Universal Robots URScript: test_first_drawing_7_m18.script

def Machining1():
  # Default parameters:
  global speed_ms = 0.3
  global speed_rads = 0.75
  global accel_mss = 3
  global accel_radss = 1.2
  global blend_radius_m = 0.001

  # Add subprograms here
  # Start of main program
  # Program generated by RoboDK v5.6.5 for UR10e on 02/02/2024 17:08:00
  # Using nominal kinematics.
  blend_radius_m = 0.001
  speed_ms = 1.000
  # set_reference(p[0.133734, -0.230000, -0.017586, 0.000000, 0.000000, 0.000000])
  set_tcp(p[0.000000, 0.000000, 0.252000, 0.000000, 0.000000, 0.000000])
  # Show Tool
  movej([-0.330517, -0.654443, -2.605811, -1.452135, 1.570796, 1.240279],accel_radss,speed_rads,0,blend_radius_m)
  movel([-0.330517, -0.654443, -2.605811, -1.452135, 1.570796, 1.240279],accel_mss,speed_ms,0,blend_radius_m)
  # Splitting Linear movement in 6 (instruction 7: MoveL 3)
  movel([-0.330517, -0.661877, -2.634190, -1.416323, 1.570796, 1.240279],accel_mss,speed_ms,0,blend_radius_m)
  movel([-0.330517, -0.671796, -2.662374, -1.378219, 1.570796, 1.240279],accel_mss,speed_ms,0,blend_radius_m)
  movel([-0.330517, -0.684615, -2.690354, -1.337420, 1.570796, 1.240279],accel_mss,speed_ms,0,blend_radius_m)
  movel([-0.330517, -0.700841, -2.718117, -1.293431, 1.570796, 1.240279],accel_mss,speed_ms,0,blend_radius_m)
  movel([-0.330517, -0.721107, -2.745644, -1.245638, 1.570796, 1.240279],accel_mss,speed_ms,0,blend_radius_m)
  movel([-0.330517, -0.746206, -2.772909, -1.193275, 1.570796, 1.240279],accel_mss,speed_ms,0,blend_radius_m)
  movel([-0.330517, -0.746206, -2.772909, -1.193275, 1.570796, 1.240279],accel_mss,speed_ms,0,blend_radius_m)
  speed_ms = 1.000
  movel([-0.330517, -0.746206, -2.772909, -1.193275, 1.570796, 1.240279],accel_mss,speed_ms,0,blend_radius_m)
  movel([-0.330517, -0.746206, -2.772909, -1.193275, 1.570796, 1.240279],accel_mss,speed_ms,0,blend_radius_m)
  movel([-0.330517, -0.746206, -2.772909, -1.193275, 1.570796, 1.240279],accel_mss,speed_ms,0,blend_radius_m)
  speed_ms = 0.005
  movel([-0.330517, -0.716695, -2.740159, -1.255535, 1.570796, 1.240279],accel_mss,speed_ms,0,blend_radius_m)
  speed_ms = 1.000
  movel([-0.330517, -0.746206, -2.772909, -1.193275, 1.570796, 1.240279],accel_mss,speed_ms,0,blend_radius_m)
  speed_ms = 0.040
  movel([-0.330517, -0.746206, -2.772909, -1.193275, 1.570796, 1.240279],accel_mss,speed_ms,0,blend_radius_m)
  speed_ms = 1.000
  movel([-0.330517, -0.746206, -2.772909, -1.193275, 1.570796, 1.240279],accel_mss,speed_ms,0,blend_radius_m)
  # Splitting Linear movement in 8 (instruction 21: MoveL 12)
  movel([-0.265752, -0.736383, -2.774388, -1.201618, 1.570796, 1.305044],accel_mss,speed_ms,0,blend_radius_m)
  movel([-0.203429, -0.731735, -2.775072, -1.205583, 1.570796, 1.367367],accel_mss,speed_ms,0,blend_radius_m)
  movel([-0.144075, -0.732399, -2.774975, -1.205016, 1.570796, 1.426722],accel_mss,speed_ms,0,blend_radius_m)
  movel([-0.088098, -0.738355, -2.774095, -1.199939, 1.570796, 1.482698],accel_mss,speed_ms,0,blend_radius_m)
  movel([-0.035774, -0.749426, -2.772413, -1.190550, 1.570796, 1.535022],accel_mss,speed_ms,0,blend_radius_m)
  movel([0.012756, -0.765294, -2.769895, -1.177200, 1.570796, 1.583552],accel_mss,speed_ms,0,blend_radius_m)
  movel([0.057475, -0.785519, -2.766498, -1.160372, 1.570796, 1.628271],accel_mss,speed_ms,0,blend_radius_m)
  movel([0.098470, -0.809577, -2.762175, -1.140637, 1.570796, 1.669266],accel_mss,speed_ms,0,blend_radius_m)
  speed_ms = 0.005
  movel([0.098470, -0.850852, -2.793539, -1.067998, 1.570796, 1.669266],accel_mss,speed_ms,0,blend_radius_m)
  speed_ms = 0.025
  movel([0.094484, -0.861595, -2.791431, -1.059363, 1.570796, 1.665281],accel_mss,speed_ms,0,blend_radius_m)
  movel([0.092287, -0.866990, -2.790348, -1.055051, 1.570796, 1.663083],accel_mss,speed_ms,0,blend_radius_m)
  movel([0.089913, -0.872383, -2.789248, -1.050758, 1.570796, 1.660710],accel_mss,speed_ms,0,blend_radius_m)
  movel([0.087338, -0.877755, -2.788135, -1.046499, 1.570796, 1.658135],accel_mss,speed_ms,0,blend_radius_m)
  movel([0.084536, -0.883089, -2.787014, -1.042286, 1.570796, 1.655333],accel_mss,speed_ms,0,blend_radius_m)
  movel([0.081477, -0.888374, -2.785886, -1.038129, 1.570796, 1.652273],accel_mss,speed_ms,0,blend_radius_m)
  movel([0.078131, -0.893592, -2.784756, -1.034042, 1.570796, 1.648928],accel_mss,speed_ms,0,blend_radius_m)
  movel([0.079373, -0.891311, -2.785252, -1.035826, 1.570796, 1.650169],accel_mss,speed_ms,0,blend_radius_m)
  movel([0.080517, -0.888452, -2.785869, -1.038068, 1.570796, 1.651313],accel_mss,speed_ms,0,blend_radius_m)
  movel([0.081210, -0.885772, -2.786443, -1.040174, 1.570796, 1.652007],accel_mss,speed_ms,0,blend_radius_m)
  movel([0.081271, -0.884745, -2.786662, -1.040982, 1.570796, 1.652068],accel_mss,speed_ms,0,blend_radius_m)
  movel([0.081086, -0.884053, -2.786809, -1.041527, 1.570796, 1.651882],accel_mss,speed_ms,0,blend_radius_m)
  movel([0.080605, -0.883776, -2.786868, -1.041745, 1.570796, 1.651401],accel_mss,speed_ms,0,blend_radius_m)
  movel([0.079917, -0.884008, -2.786819, -1.041563, 1.570796, 1.650713],accel_mss,speed_ms,0,blend_radius_m)
  movel([0.079063, -0.884679, -2.786676, -1.041034, 1.570796, 1.649859],accel_mss,speed_ms,0,blend_radius_m)
  movel([0.078060, -0.885737, -2.786451, -1.040201, 1.570796, 1.648856],accel_mss,speed_ms,0,blend_radius_m)
  movel([0.075754, -0.888735, -2.785808, -1.037846, 1.570796, 1.646551],accel_mss,speed_ms,0,blend_radius_m)
  movel([0.073242, -0.892488, -2.784996, -1.034905, 1.570796, 1.644038],accel_mss,speed_ms,0,blend_radius_m)
  movel([0.068514, -0.900288, -2.783281, -1.028820, 1.570796, 1.639311],accel_mss,speed_ms,0,blend_radius_m)
  movel([0.065663, -0.905241, -2.782172, -1.024976, 1.570796, 1.636460],accel_mss,speed_ms,0,blend_radius_m)
  movel([0.061416, -0.912163, -2.780598, -1.019629, 1.570796, 1.632212],accel_mss,speed_ms,0,blend_radius_m)
  movel([0.059067, -0.915476, -2.779833, -1.017080, 1.570796, 1.629863],accel_mss,speed_ms,0,blend_radius_m)
  movel([0.056470, -0.918581, -2.779110, -1.014698, 1.570796, 1.627267],accel_mss,speed_ms,0,blend_radius_m)
  movel([0.057008, -0.917651, -2.779327, -1.015410, 1.570796, 1.627804],accel_mss,speed_ms,0,blend_radius_m)
  movel([0.057386, -0.916311, -2.779639, -1.016439, 1.570796, 1.628182],accel_mss,speed_ms,0,blend_radius_m)
  movel([0.057710, -0.913007, -2.780403, -1.018979, 1.570796, 1.628506],accel_mss,speed_ms,0,blend_radius_m)
  movel([0.057532, -0.909923, -2.781110, -1.021356, 1.570796, 1.628328],accel_mss,speed_ms,0,blend_radius_m)
  movel([0.057276, -0.908855, -2.781354, -1.022180, 1.570796, 1.628072],accel_mss,speed_ms,0,blend_radius_m)
  movel([0.056930, -0.908319, -2.781476, -1.022594, 1.570796, 1.627726],accel_mss,speed_ms,0,blend_radius_m)
  movel([0.055907, -0.908068, -2.781533, -1.022788, 1.570796, 1.626704],accel_mss,speed_ms,0,blend_radius_m)
  movel([0.054873, -0.908367, -2.781465, -1.022557, 1.570796, 1.625669],accel_mss,speed_ms,0,blend_radius_m)
  movel([0.053834, -0.909106, -2.781297, -1.021987, 1.570796, 1.624631],accel_mss,speed_ms,0,blend_radius_m)
  movel([0.052803, -0.910180, -2.781052, -1.021157, 1.570796, 1.623599],accel_mss,speed_ms,0,blend_radius_m)
  movel([0.050825, -0.912852, -2.780439, -1.019098, 1.570796, 1.621621],accel_mss,speed_ms,0,blend_radius_m)
  movel([0.049035, -0.915498, -2.779828, -1.017063, 1.570796, 1.619831],accel_mss,speed_ms,0,blend_radius_m)
  movel([0.046096, -0.919482, -2.778899, -1.014007, 1.570796, 1.616892],accel_mss,speed_ms,0,blend_radius_m)
  movel([0.043104, -0.923120, -2.778043, -1.011226, 1.570796, 1.613900],accel_mss,speed_ms,0,blend_radius_m)
  movel([0.039882, -0.926413, -2.777260, -1.008716, 1.570796, 1.610679],accel_mss,speed_ms,0,blend_radius_m)
  movel([0.036270, -0.929334, -2.776560, -1.006495, 1.570796, 1.607066],accel_mss,speed_ms,0,blend_radius_m)
  movel([0.038295, -0.926302, -2.777286, -1.008800, 1.570796, 1.609092],accel_mss,speed_ms,0,blend_radius_m)
  movel([0.039935, -0.923235, -2.778015, -1.011138, 1.570796, 1.610731],accel_mss,speed_ms,0,blend_radius_m)
  movel([0.040448, -0.921718, -2.778374, -1.012297, 1.570796, 1.611244],accel_mss,speed_ms,0,blend_radius_m)
  movel([0.040644, -0.920343, -2.778697, -1.013349, 1.570796, 1.611440],accel_mss,speed_ms,0,blend_radius_m)
  movel([0.040480, -0.919233, -2.778958, -1.014198, 1.570796, 1.611276],accel_mss,speed_ms,0,blend_radius_m)
  movel([0.039889, -0.918538, -2.779120, -1.014731, 1.570796, 1.610686],accel_mss,speed_ms,0,blend_radius_m)
  movel([0.038611, -0.918412, -2.779150, -1.014827, 1.570796, 1.609407],accel_mss,speed_ms,0,blend_radius_m)
  movel([0.036998, -0.918988, -2.779015, -1.014386, 1.570796, 1.607794],accel_mss,speed_ms,0,blend_radius_m)
  movel([0.035210, -0.920033, -2.778770, -1.013586, 1.570796, 1.606006],accel_mss,speed_ms,0,blend_radius_m)
  movel([0.033415, -0.921289, -2.778475, -1.012625, 1.570796, 1.604211],accel_mss,speed_ms,0,blend_radius_m)
  speed_ms = 0.005
  movel([0.033415, -0.911749, -2.772496, -1.028143, 1.570796, 1.604211],accel_mss,speed_ms,0,blend_radius_m)
  speed_ms = 0.040
  movel([0.037572, -0.944814, -2.764429, -1.003146, 1.570796, 1.608368],accel_mss,speed_ms,0,blend_radius_m)
  speed_ms = 0.005
  movel([0.037572, -0.954534, -2.770284, -0.987571, 1.570796, 1.608368],accel_mss,speed_ms,0,blend_radius_m)
  speed_ms = 0.025
  movel([0.038407, -0.952070, -2.770916, -0.989403, 1.570796, 1.609204],accel_mss,speed_ms,0,blend_radius_m)
  movel([0.039504, -0.949536, -2.771562, -0.991291, 1.570796, 1.610300],accel_mss,speed_ms,0,blend_radius_m)
  movel([0.040832, -0.946976, -2.772211, -0.993202, 1.570796, 1.611628],accel_mss,speed_ms,0,blend_radius_m)
  movel([0.042377, -0.944420, -2.772854, -0.995116, 1.570796, 1.613173],accel_mss,speed_ms,0,blend_radius_m)
  movel([0.044112, -0.941903, -2.773482, -0.997004, 1.570796, 1.614908],accel_mss,speed_ms,0,blend_radius_m)
  movel([0.046017, -0.939467, -2.774087, -0.998835, 1.570796, 1.616813],accel_mss,speed_ms,0,blend_radius_m)
  movel([0.048065, -0.937149, -2.774659, -1.000582, 1.570796, 1.618862],accel_mss,speed_ms,0,blend_radius_m)
  movel([0.050239, -0.934981, -2.775190, -1.002218, 1.570796, 1.621035],accel_mss,speed_ms,0,blend_radius_m)
  movel([0.053602, -0.932102, -2.775891, -1.004396, 1.570796, 1.624398],accel_mss,speed_ms,0,blend_radius_m)
  movel([0.056890, -0.929797, -2.776448, -1.006144, 1.570796, 1.627686],accel_mss,speed_ms,0,blend_radius_m)
  movel([0.060092, -0.928029, -2.776873, -1.007487, 1.570796, 1.630888],accel_mss,speed_ms,0,blend_radius_m)
  movel([0.063188, -0.926767, -2.777175, -1.008446, 1.570796, 1.633984],accel_mss,speed_ms,0,blend_radius_m)
  movel([0.066168, -0.925977, -2.777364, -1.009048, 1.570796, 1.636964],accel_mss,speed_ms,0,blend_radius_m)
  movel([0.069022, -0.925620, -2.777449, -1.009320, 1.570796, 1.639818],accel_mss,speed_ms,0,blend_radius_m)
  movel([0.071734, -0.925666, -2.777438, -1.009285, 1.570796, 1.642530],accel_mss,speed_ms,0,blend_radius_m)
  movel([0.074296, -0.926070, -2.777342, -1.008977, 1.570796, 1.645092],accel_mss,speed_ms,0,blend_radius_m)
  movel([0.076697, -0.926796, -2.777168, -1.008425, 1.570796, 1.647493],accel_mss,speed_ms,0,blend_radius_m)
  movel([0.078931, -0.927802, -2.776927, -1.007659, 1.570796, 1.649727],accel_mss,speed_ms,0,blend_radius_m)
  movel([0.082865, -0.930490, -2.776281, -1.005618, 1.570796, 1.653661],accel_mss,speed_ms,0,blend_radius_m)
  movel([0.086044, -0.933794, -2.775479, -1.003115, 1.570796, 1.656840],accel_mss,speed_ms,0,blend_radius_m)
  movel([0.088410, -0.937397, -2.774597, -1.000394, 1.570796, 1.659206],accel_mss,speed_ms,0,blend_radius_m)
  movel([0.090331, -0.941611, -2.773555, -0.997223, 1.570796, 1.661127],accel_mss,speed_ms,0,blend_radius_m)
  movel([0.091833, -0.946185, -2.772410, -0.993794, 1.570796, 1.662629],accel_mss,speed_ms,0,blend_radius_m)
  movel([0.092966, -0.951056, -2.771175, -0.990158, 1.570796, 1.663762],accel_mss,speed_ms,0,blend_radius_m)
  movel([0.093774, -0.956168, -2.769862, -0.986359, 1.570796, 1.664570],accel_mss,speed_ms,0,blend_radius_m)
  movel([0.094306, -0.961464, -2.768483, -0.982443, 1.570796, 1.665103],accel_mss,speed_ms,0,blend_radius_m)
  movel([0.094614, -0.966887, -2.767050, -0.978453, 1.570796, 1.665411],accel_mss,speed_ms,0,blend_radius_m)
  movel([0.094736, -0.977899, -2.764077, -0.970413, 1.570796, 1.665532],accel_mss,speed_ms,0,blend_radius_m)
  movel([0.094750, -0.985564, -2.761956, -0.964869, 1.570796, 1.665546],accel_mss,speed_ms,0,blend_radius_m)
  movel([0.095064, -0.989150, -2.760950, -0.962290, 1.570796, 1.665861],accel_mss,speed_ms,0,blend_radius_m)
  movel([0.095787, -0.992414, -2.760025, -0.959950, 1.570796, 1.666583],accel_mss,speed_ms,0,blend_radius_m)
  movel([0.097346, -0.996214, -2.758939, -0.957236, 1.570796, 1.668143],accel_mss,speed_ms,0,blend_radius_m)
  movel([0.098905, -1.000023, -2.757839, -0.954527, 1.570796, 1.669701],accel_mss,speed_ms,0,blend_radius_m)
  movel([0.099406, -1.002068, -2.757244, -0.953076, 1.570796, 1.670202],accel_mss,speed_ms,0,blend_radius_m)
  movel([0.099571, -1.004282, -2.756597, -0.951510, 1.570796, 1.670367],accel_mss,speed_ms,0,blend_radius_m)
  movel([0.099295, -1.006711, -2.755882, -0.949796, 1.570796, 1.670091],accel_mss,speed_ms,0,blend_radius_m)
  movel([0.098473, -1.009410, -2.755083, -0.947896, 1.570796, 1.669269],accel_mss,speed_ms,0,blend_radius_m)
  movel([0.101094, -1.002602, -2.757088, -0.952698, 1.570796, 1.671890],accel_mss,speed_ms,0,blend_radius_m)
  movel([0.103419, -0.995838, -2.759047, -0.957504, 1.570796, 1.674215],accel_mss,speed_ms,0,blend_radius_m)
  movel([0.107547, -0.982266, -2.762874, -0.967249, 1.570796, 1.678343],accel_mss,speed_ms,0,blend_radius_m)
  movel([0.109649, -0.974669, -2.764958, -0.972762, 1.570796, 1.680446],accel_mss,speed_ms,0,blend_radius_m)
  movel([0.111578, -0.967069, -2.767001, -0.978319, 1.570796, 1.682375],accel_mss,speed_ms,0,blend_radius_m)
  movel([0.115043, -0.951807, -2.770983, -0.989598, 1.570796, 1.685839],accel_mss,speed_ms,0,blend_radius_m)
  movel([0.118016, -0.936784, -2.774748, -1.000856, 1.570796, 1.688812],accel_mss,speed_ms,0,blend_radius_m)
  movel([0.119175, -0.929313, -2.776564, -1.006511, 1.570796, 1.689972],accel_mss,speed_ms,0,blend_radius_m)
  movel([0.119952, -0.922044, -2.778297, -1.012048, 1.570796, 1.690749],accel_mss,speed_ms,0,blend_radius_m)
  movel([0.120167, -0.916526, -2.779589, -1.016273, 1.570796, 1.690963],accel_mss,speed_ms,0,blend_radius_m)
  movel([0.120127, -0.911118, -2.780837, -1.020434, 1.570796, 1.690923],accel_mss,speed_ms,0,blend_radius_m)
  movel([0.120107, -0.905634, -2.782084, -1.024671, 1.570796, 1.690904],accel_mss,speed_ms,0,blend_radius_m)
  movel([0.120387, -0.899887, -2.783370, -1.029132, 1.570796, 1.691183],accel_mss,speed_ms,0,blend_radius_m)
  movel([0.120647, -0.898247, -2.783733, -1.030409, 1.570796, 1.691443],accel_mss,speed_ms,0,blend_radius_m)
  movel([0.121203, -0.896466, -2.784126, -1.031797, 1.570796, 1.692000],accel_mss,speed_ms,0,blend_radius_m)
  movel([0.122110, -0.894787, -2.784494, -1.033107, 1.570796, 1.692906],accel_mss,speed_ms,0,blend_radius_m)
  movel([0.122719, -0.894054, -2.784655, -1.033680, 1.570796, 1.693515],accel_mss,speed_ms,0,blend_radius_m)
  movel([0.123441, -0.893428, -2.784791, -1.034169, 1.570796, 1.694238],accel_mss,speed_ms,0,blend_radius_m)
  movel([0.124465, -0.892889, -2.784909, -1.034591, 1.570796, 1.695262],accel_mss,speed_ms,0,blend_radius_m)
  movel([0.125422, -0.892628, -2.784965, -1.034795, 1.570796, 1.696219],accel_mss,speed_ms,0,blend_radius_m)
  movel([0.130425, -0.891913, -2.785121, -1.035355, 1.570796, 1.701221],accel_mss,speed_ms,0,blend_radius_m)
  movel([0.134885, -0.891965, -2.785110, -1.035315, 1.570796, 1.705681],accel_mss,speed_ms,0,blend_radius_m)
  movel([0.138838, -0.892713, -2.784947, -1.034729, 1.570796, 1.709634],accel_mss,speed_ms,0,blend_radius_m)
  movel([0.142320, -0.894105, -2.784643, -1.033640, 1.570796, 1.713117],accel_mss,speed_ms,0,blend_radius_m)
  movel([0.145368, -0.896070, -2.784213, -1.032106, 1.570796, 1.716164],accel_mss,speed_ms,0,blend_radius_m)
  movel([0.148021, -0.898542, -2.783668, -1.030179, 1.570796, 1.718817],accel_mss,speed_ms,0,blend_radius_m)
  movel([0.150317, -0.901457, -2.783021, -1.027911, 1.570796, 1.721113],accel_mss,speed_ms,0,blend_radius_m)
  movel([0.152293, -0.904755, -2.782282, -1.025352, 1.570796, 1.723089],accel_mss,speed_ms,0,blend_radius_m)
  movel([0.153993, -0.908367, -2.781465, -1.022557, 1.570796, 1.724789],accel_mss,speed_ms,0,blend_radius_m)
  movel([0.155459, -0.912228, -2.780583, -1.019578, 1.570796, 1.726255],accel_mss,speed_ms,0,blend_radius_m)
  movel([0.157842, -0.920452, -2.778672, -1.013265, 1.570796, 1.728639],accel_mss,speed_ms,0,blend_radius_m)
  movel([0.161526, -0.937276, -2.774627, -1.000486, 1.570796, 1.732322],accel_mss,speed_ms,0,blend_radius_m)
  movel([0.162250, -0.939773, -2.774011, -0.998605, 1.570796, 1.733046],accel_mss,speed_ms,0,blend_radius_m)
  movel([0.162856, -0.940764, -2.773765, -0.997859, 1.570796, 1.733653],accel_mss,speed_ms,0,blend_radius_m)
  movel([0.163731, -0.941443, -2.773597, -0.997349, 1.570796, 1.734527],accel_mss,speed_ms,0,blend_radius_m)
  movel([0.165528, -0.941709, -2.773531, -0.997150, 1.570796, 1.736325],accel_mss,speed_ms,0,blend_radius_m)
  movel([0.166517, -0.941509, -2.773580, -0.997300, 1.570796, 1.737313],accel_mss,speed_ms,0,blend_radius_m)
  movel([0.167553, -0.941108, -2.773680, -0.997601, 1.570796, 1.738350],accel_mss,speed_ms,0,blend_radius_m)
  movel([0.169715, -0.939801, -2.774004, -0.998584, 1.570796, 1.740512],accel_mss,speed_ms,0,blend_radius_m)
  movel([0.171931, -0.937949, -2.774462, -0.999978, 1.570796, 1.742727],accel_mss,speed_ms,0,blend_radius_m)
  movel([0.174106, -0.935721, -2.775009, -1.001659, 1.570796, 1.744902],accel_mss,speed_ms,0,blend_radius_m)
  movel([0.176150, -0.933279, -2.775605, -1.003505, 1.570796, 1.746946],accel_mss,speed_ms,0,blend_radius_m)
  movel([0.177974, -0.930783, -2.776210, -1.005396, 1.570796, 1.748770],accel_mss,speed_ms,0,blend_radius_m)
  movel([0.179471, -0.928409, -2.776782, -1.007198, 1.570796, 1.750268],accel_mss,speed_ms,0,blend_radius_m)
  movel([0.181767, -0.924306, -2.777762, -1.010321, 1.570796, 1.752563],accel_mss,speed_ms,0,blend_radius_m)
  movel([0.183931, -0.920150, -2.778743, -1.013496, 1.570796, 1.754728],accel_mss,speed_ms,0,blend_radius_m)
  movel([0.187846, -0.911748, -2.780693, -1.019948, 1.570796, 1.758643],accel_mss,speed_ms,0,blend_radius_m)
  movel([0.191204, -0.903342, -2.782599, -1.026448, 1.570796, 1.762001],accel_mss,speed_ms,0,blend_radius_m)
  movel([0.193979, -0.895073, -2.784432, -1.032884, 1.570796, 1.764775],accel_mss,speed_ms,0,blend_radius_m)
  movel([0.194923, -0.891979, -2.785107, -1.035303, 1.570796, 1.765719],accel_mss,speed_ms,0,blend_radius_m)
  movel([0.196094, -0.888834, -2.785787, -1.037769, 1.570796, 1.766891],accel_mss,speed_ms,0,blend_radius_m)
  movel([0.196862, -0.887263, -2.786124, -1.039002, 1.570796, 1.767658],accel_mss,speed_ms,0,blend_radius_m)
  movel([0.197803, -0.885695, -2.786460, -1.040235, 1.570796, 1.768600],accel_mss,speed_ms,0,blend_radius_m)
  movel([0.198955, -0.884142, -2.786790, -1.041457, 1.570796, 1.769752],accel_mss,speed_ms,0,blend_radius_m)
  movel([0.200357, -0.882615, -2.787114, -1.042660, 1.570796, 1.771153],accel_mss,speed_ms,0,blend_radius_m)
  movel([0.202401, -0.881008, -2.787453, -1.043928, 1.570796, 1.773197],accel_mss,speed_ms,0,blend_radius_m)
  movel([0.204401, -0.880128, -2.787638, -1.044623, 1.570796, 1.775198],accel_mss,speed_ms,0,blend_radius_m)
  movel([0.206224, -0.879892, -2.787688, -1.044809, 1.570796, 1.777021],accel_mss,speed_ms,0,blend_radius_m)
  movel([0.207752, -0.880207, -2.787622, -1.044560, 1.570796, 1.778548],accel_mss,speed_ms,0,blend_radius_m)
  movel([0.209849, -0.881389, -2.787373, -1.043627, 1.570796, 1.780645],accel_mss,speed_ms,0,blend_radius_m)
  movel([0.211668, -0.882983, -2.787036, -1.042370, 1.570796, 1.782464],accel_mss,speed_ms,0,blend_radius_m)
  movel([0.214678, -0.886847, -2.786213, -1.039329, 1.570796, 1.785474],accel_mss,speed_ms,0,blend_radius_m)
  movel([0.215840, -0.888920, -2.785768, -1.037701, 1.570796, 1.786637],accel_mss,speed_ms,0,blend_radius_m)
  movel([0.216722, -0.891180, -2.785280, -1.035929, 1.570796, 1.787518],accel_mss,speed_ms,0,blend_radius_m)
  movel([0.217344, -0.893608, -2.784752, -1.034029, 1.570796, 1.788140],accel_mss,speed_ms,0,blend_radius_m)
  movel([0.217717, -0.896195, -2.784185, -1.032008, 1.570796, 1.788513],accel_mss,speed_ms,0,blend_radius_m)
  movel([0.217858, -0.898923, -2.783584, -1.029882, 1.570796, 1.788654],accel_mss,speed_ms,0,blend_radius_m)
  movel([0.217499, -0.904763, -2.782280, -1.025346, 1.570796, 1.788295],accel_mss,speed_ms,0,blend_radius_m)
  movel([0.217027, -0.907846, -2.781583, -1.022960, 1.570796, 1.787823],accel_mss,speed_ms,0,blend_radius_m)
  movel([0.215585, -0.914270, -2.780112, -1.018007, 1.570796, 1.786381],accel_mss,speed_ms,0,blend_radius_m)
  movel([0.213564, -0.920962, -2.778552, -1.012875, 1.570796, 1.784360],accel_mss,speed_ms,0,blend_radius_m)
  movel([0.211074, -0.927836, -2.776919, -1.007633, 1.570796, 1.781870],accel_mss,speed_ms,0,blend_radius_m)
  movel([0.208233, -0.934789, -2.775237, -1.002363, 1.570796, 1.779029],accel_mss,speed_ms,0,blend_radius_m)
  movel([0.203631, -0.944939, -2.772723, -0.994727, 1.570796, 1.774427],accel_mss,speed_ms,0,blend_radius_m)
  movel([0.201108, -0.949995, -2.771446, -0.990948, 1.570796, 1.771904],accel_mss,speed_ms,0,blend_radius_m)
  movel([0.198410, -0.955010, -2.770161, -0.987218, 1.570796, 1.769207],accel_mss,speed_ms,0,blend_radius_m)
  movel([0.195524, -0.959954, -2.768878, -0.983557, 1.570796, 1.766320],accel_mss,speed_ms,0,blend_radius_m)
  movel([0.192436, -0.964804, -2.767603, -0.979982, 1.570796, 1.763232],accel_mss,speed_ms,0,blend_radius_m)
  movel([0.189119, -0.969547, -2.766339, -0.976502, 1.570796, 1.759915],accel_mss,speed_ms,0,blend_radius_m)
  movel([0.185564, -0.974153, -2.765098, -0.973139, 1.570796, 1.756360],accel_mss,speed_ms,0,blend_radius_m)
  movel([0.180277, -0.980341, -2.763406, -0.968642, 1.570796, 1.751073],accel_mss,speed_ms,0,blend_radius_m)
  movel([0.177371, -0.983434, -2.762550, -0.966406, 1.570796, 1.748167],accel_mss,speed_ms,0,blend_radius_m)
  movel([0.174357, -0.986357, -2.761734, -0.964297, 1.570796, 1.745154],accel_mss,speed_ms,0,blend_radius_m)
  movel([0.171294, -0.988986, -2.760996, -0.962407, 1.570796, 1.742090],accel_mss,speed_ms,0,blend_radius_m)
  movel([0.168232, -0.991197, -2.760371, -0.960822, 1.570796, 1.739028],accel_mss,speed_ms,0,blend_radius_m)
  movel([0.165220, -0.992864, -2.759897, -0.959628, 1.570796, 1.736016],accel_mss,speed_ms,0,blend_radius_m)
  movel([0.163750, -0.993460, -2.759727, -0.959202, 1.570796, 1.734546],accel_mss,speed_ms,0,blend_radius_m)
  movel([0.162314, -0.993869, -2.759610, -0.958910, 1.570796, 1.733110],accel_mss,speed_ms,0,blend_radius_m)
  movel([0.160767, -0.994093, -2.759546, -0.958749, 1.570796, 1.731564],accel_mss,speed_ms,0,blend_radius_m)
  movel([0.159366, -0.994058, -2.759556, -0.958774, 1.570796, 1.730163],accel_mss,speed_ms,0,blend_radius_m)
  movel([0.158098, -0.993791, -2.759633, -0.958966, 1.570796, 1.728894],accel_mss,speed_ms,0,blend_radius_m)
  movel([0.156956, -0.993308, -2.759770, -0.959311, 1.570796, 1.727752],accel_mss,speed_ms,0,blend_radius_m)
  movel([0.155007, -0.991802, -2.760199, -0.960388, 1.570796, 1.725804],accel_mss,speed_ms,0,blend_radius_m)
  movel([0.153455, -0.989715, -2.760790, -0.961884, 1.570796, 1.724251],accel_mss,speed_ms,0,blend_radius_m)
  movel([0.152226, -0.987238, -2.761488, -0.963664, 1.570796, 1.723022],accel_mss,speed_ms,0,blend_radius_m)
  movel([0.151254, -0.984552, -2.762239, -0.965599, 1.570796, 1.722051],accel_mss,speed_ms,0,blend_radius_m)
  movel([0.149812, -0.979297, -2.763693, -0.969399, 1.570796, 1.720608],accel_mss,speed_ms,0,blend_radius_m)
  movel([0.149169, -0.976821, -2.764372, -0.971196, 1.570796, 1.719965],accel_mss,speed_ms,0,blend_radius_m)
  movel([0.148254, -0.974605, -2.764975, -0.972809, 1.570796, 1.719050],accel_mss,speed_ms,0,blend_radius_m)
  movel([0.147575, -0.973756, -2.765205, -0.973427, 1.570796, 1.718371],accel_mss,speed_ms,0,blend_radius_m)
  movel([0.146683, -0.973163, -2.765366, -0.973860, 1.570796, 1.717479],accel_mss,speed_ms,0,blend_radius_m)
  movel([0.145535, -0.972893, -2.765439, -0.974057, 1.570796, 1.716332],accel_mss,speed_ms,0,blend_radius_m)
  movel([0.144083, -0.973006, -2.765408, -0.973975, 1.570796, 1.714879],accel_mss,speed_ms,0,blend_radius_m)
  movel([0.144394, -0.973052, -2.765396, -0.973941, 1.570796, 1.715191],accel_mss,speed_ms,0,blend_radius_m)
  movel([0.144561, -0.973335, -2.765319, -0.973734, 1.570796, 1.715357],accel_mss,speed_ms,0,blend_radius_m)
  movel([0.144480, -0.974556, -2.764988, -0.972845, 1.570796, 1.715276],accel_mss,speed_ms,0,blend_radius_m)
  movel([0.143903, -0.976547, -2.764446, -0.971395, 1.570796, 1.714700],accel_mss,speed_ms,0,blend_radius_m)
  movel([0.142911, -0.979182, -2.763725, -0.969482, 1.570796, 1.713708],accel_mss,speed_ms,0,blend_radius_m)
  movel([0.139967, -0.985880, -2.761868, -0.964641, 1.570796, 1.710763],accel_mss,speed_ms,0,blend_radius_m)
  movel([0.136215, -0.993659, -2.759670, -0.959059, 1.570796, 1.707011],accel_mss,speed_ms,0,blend_radius_m)
  movel([0.128486, -1.008701, -2.755293, -0.948395, 1.570796, 1.699282],accel_mss,speed_ms,0,blend_radius_m)
  movel([0.123866, -1.017165, -2.752755, -0.942469, 1.570796, 1.694663],accel_mss,speed_ms,0,blend_radius_m)
  movel([0.118500, -1.025835, -2.750097, -0.936457, 1.570796, 1.689296],accel_mss,speed_ms,0,blend_radius_m)
  movel([0.113088, -1.034273, -2.747454, -0.930662, 1.570796, 1.683885],accel_mss,speed_ms,0,blend_radius_m)
  movel([0.107607, -1.042564, -2.744801, -0.925024, 1.570796, 1.678403],accel_mss,speed_ms,0,blend_radius_m)
  movel([0.096784, -1.058318, -2.739605, -0.914466, 1.570796, 1.667580],accel_mss,speed_ms,0,blend_radius_m)
  movel([0.091340, -1.065635, -2.737121, -0.909633, 1.570796, 1.662136],accel_mss,speed_ms,0,blend_radius_m)
  movel([0.088492, -1.069136, -2.735917, -0.907336, 1.570796, 1.659288],accel_mss,speed_ms,0,blend_radius_m)
  movel([0.085541, -1.072496, -2.734751, -0.905142, 1.570796, 1.656337],accel_mss,speed_ms,0,blend_radius_m)
  movel([0.082458, -1.075684, -2.733635, -0.903069, 1.570796, 1.653255],accel_mss,speed_ms,0,blend_radius_m)
  movel([0.079236, -1.078673, -2.732582, -0.901134, 1.570796, 1.650032],accel_mss,speed_ms,0,blend_radius_m)
  movel([0.080076, -1.072663, -2.734693, -0.905033, 1.570796, 1.650872],accel_mss,speed_ms,0,blend_radius_m)
  movel([0.080087, -1.070990, -2.735275, -0.906125, 1.570796, 1.650884],accel_mss,speed_ms,0,blend_radius_m)
  movel([0.079804, -1.070415, -2.735474, -0.906500, 1.570796, 1.650600],accel_mss,speed_ms,0,blend_radius_m)
  movel([0.079211, -1.070213, -2.735544, -0.906632, 1.570796, 1.650008],accel_mss,speed_ms,0,blend_radius_m)
  movel([0.078545, -1.070393, -2.735482, -0.906514, 1.570796, 1.649341],accel_mss,speed_ms,0,blend_radius_m)
  movel([0.077831, -1.070816, -2.735335, -0.906238, 1.570796, 1.648627],accel_mss,speed_ms,0,blend_radius_m)
  movel([0.074420, -1.073503, -2.734399, -0.904486, 1.570796, 1.645216],accel_mss,speed_ms,0,blend_radius_m)
  movel([0.072411, -1.074760, -2.733960, -0.903669, 1.570796, 1.643207],accel_mss,speed_ms,0,blend_radius_m)
  movel([0.070406, -1.075731, -2.733619, -0.903039, 1.570796, 1.641202],accel_mss,speed_ms,0,blend_radius_m)
  movel([0.068457, -1.076392, -2.733387, -0.902610, 1.570796, 1.639253],accel_mss,speed_ms,0,blend_radius_m)
  movel([0.067876, -1.076424, -2.733376, -0.902590, 1.570796, 1.638673],accel_mss,speed_ms,0,blend_radius_m)
  movel([0.067717, -1.076086, -2.733494, -0.902809, 1.570796, 1.638514],accel_mss,speed_ms,0,blend_radius_m)
  movel([0.068293, -1.074277, -2.734129, -0.903983, 1.570796, 1.639089],accel_mss,speed_ms,0,blend_radius_m)
  movel([0.068248, -1.073755, -2.734312, -0.904323, 1.570796, 1.639044],accel_mss,speed_ms,0,blend_radius_m)
  movel([0.067937, -1.073447, -2.734419, -0.904523, 1.570796, 1.638733],accel_mss,speed_ms,0,blend_radius_m)
  movel([0.067444, -1.073351, -2.734453, -0.904586, 1.570796, 1.638240],accel_mss,speed_ms,0,blend_radius_m)
  movel([0.066848, -1.073466, -2.734412, -0.904511, 1.570796, 1.637644],accel_mss,speed_ms,0,blend_radius_m)
  movel([0.065582, -1.074163, -2.734169, -0.904057, 1.570796, 1.636378],accel_mss,speed_ms,0,blend_radius_m)
  movel([0.056656, -1.081474, -2.731587, -0.899328, 1.570796, 1.627452],accel_mss,speed_ms,0,blend_radius_m)
  movel([0.059293, -1.078836, -2.732524, -0.901029, 1.570796, 1.630089],accel_mss,speed_ms,0,blend_radius_m)
  movel([0.061894, -1.075999, -2.733525, -0.902865, 1.570796, 1.632691],accel_mss,speed_ms,0,blend_radius_m)
  movel([0.064438, -1.073011, -2.734571, -0.904807, 1.570796, 1.635234],accel_mss,speed_ms,0,blend_radius_m)
  movel([0.066915, -1.069903, -2.735651, -0.906834, 1.570796, 1.637712],accel_mss,speed_ms,0,blend_radius_m)
  movel([0.071603, -1.063485, -2.737856, -0.911048, 1.570796, 1.642399],accel_mss,speed_ms,0,blend_radius_m)
  movel([0.075821, -1.057076, -2.740022, -0.915291, 1.570796, 1.646617],accel_mss,speed_ms,0,blend_radius_m)
  movel([0.080132, -1.050034, -2.742363, -0.919992, 1.570796, 1.650928],accel_mss,speed_ms,0,blend_radius_m)
  movel([0.084250, -1.042837, -2.744713, -0.924839, 1.570796, 1.655047],accel_mss,speed_ms,0,blend_radius_m)
  movel([0.086168, -1.039200, -2.745884, -0.927305, 1.570796, 1.656965],accel_mss,speed_ms,0,blend_radius_m)
  movel([0.087963, -1.035546, -2.747050, -0.929793, 1.570796, 1.658760],accel_mss,speed_ms,0,blend_radius_m)
  movel([0.089601, -1.031889, -2.748206, -0.932293, 1.570796, 1.660397],accel_mss,speed_ms,0,blend_radius_m)
  movel([0.091057, -1.028231, -2.749352, -0.934805, 1.570796, 1.661853],accel_mss,speed_ms,0,blend_radius_m)
  movel([0.091816, -1.025973, -2.750054, -0.936361, 1.570796, 1.662613],accel_mss,speed_ms,0,blend_radius_m)
  movel([0.092410, -1.023740, -2.750745, -0.937904, 1.570796, 1.663206],accel_mss,speed_ms,0,blend_radius_m)
  movel([0.093141, -1.019370, -2.752085, -0.940935, 1.570796, 1.663937],accel_mss,speed_ms,0,blend_radius_m)
  movel([0.093305, -1.015177, -2.753356, -0.943856, 1.570796, 1.664101],accel_mss,speed_ms,0,blend_radius_m)
  movel([0.092955, -1.011216, -2.754545, -0.946628, 1.570796, 1.663751],accel_mss,speed_ms,0,blend_radius_m)
  movel([0.092159, -1.007532, -2.755640, -0.949217, 1.570796, 1.662955],accel_mss,speed_ms,0,blend_radius_m)
  movel([0.090980, -1.004179, -2.756627, -0.951583, 1.570796, 1.661776],accel_mss,speed_ms,0,blend_radius_m)
  movel([0.089473, -1.001211, -2.757494, -0.953684, 1.570796, 1.660269],accel_mss,speed_ms,0,blend_radius_m)
  movel([0.087711, -0.998675, -2.758230, -0.955485, 1.570796, 1.658507],accel_mss,speed_ms,0,blend_radius_m)
  movel([0.086357, -0.997636, -2.758530, -0.956223, 1.570796, 1.657154],accel_mss,speed_ms,0,blend_radius_m)
  movel([0.084665, -0.997306, -2.758625, -0.956458, 1.570796, 1.655461],accel_mss,speed_ms,0,blend_radius_m)
  movel([0.082738, -0.997630, -2.758531, -0.956228, 1.570796, 1.653534],accel_mss,speed_ms,0,blend_radius_m)
  movel([0.080685, -0.998552, -2.758265, -0.955572, 1.570796, 1.651481],accel_mss,speed_ms,0,blend_radius_m)
  movel([0.078604, -1.000010, -2.757843, -0.954536, 1.570796, 1.649400],accel_mss,speed_ms,0,blend_radius_m)
  movel([0.076600, -1.001946, -2.757280, -0.953163, 1.570796, 1.647396],accel_mss,speed_ms,0,blend_radius_m)
  movel([0.074785, -1.004292, -2.756594, -0.951503, 1.570796, 1.645582],accel_mss,speed_ms,0,blend_radius_m)
  movel([0.073255, -1.006987, -2.755801, -0.949601, 1.570796, 1.644052],accel_mss,speed_ms,0,blend_radius_m)
  movel([0.071220, -1.011114, -2.754575, -0.946700, 1.570796, 1.642016],accel_mss,speed_ms,0,blend_radius_m)
  movel([0.069032, -1.015194, -2.753351, -0.943844, 1.570796, 1.639828],accel_mss,speed_ms,0,blend_radius_m)
  movel([0.066672, -1.019192, -2.752139, -0.941058, 1.570796, 1.637469],accel_mss,speed_ms,0,blend_radius_m)
  movel([0.064115, -1.023085, -2.750947, -0.938357, 1.570796, 1.634912],accel_mss,speed_ms,0,blend_radius_m)
  movel([0.061349, -1.026837, -2.749786, -0.935766, 1.570796, 1.632145],accel_mss,speed_ms,0,blend_radius_m)
  movel([0.058346, -1.030424, -2.748667, -0.933299, 1.570796, 1.629142],accel_mss,speed_ms,0,blend_radius_m)
  movel([0.055086, -1.033820, -2.747597, -0.930972, 1.570796, 1.625883],accel_mss,speed_ms,0,blend_radius_m)
  movel([0.051553, -1.036996, -2.746589, -0.928805, 1.570796, 1.622350],accel_mss,speed_ms,0,blend_radius_m)
  movel([0.049638, -1.038441, -2.746127, -0.927821, 1.570796, 1.620435],accel_mss,speed_ms,0,blend_radius_m)
  movel([0.047695, -1.039662, -2.745736, -0.926991, 1.570796, 1.618491],accel_mss,speed_ms,0,blend_radius_m)
  movel([0.043791, -1.041691, -2.745083, -0.925615, 1.570796, 1.614588],accel_mss,speed_ms,0,blend_radius_m)
  movel([0.040756, -1.042978, -2.744667, -0.924744, 1.570796, 1.611552],accel_mss,speed_ms,0,blend_radius_m)
  movel([0.037886, -1.043831, -2.744391, -0.924167, 1.570796, 1.608683],accel_mss,speed_ms,0,blend_radius_m)
  movel([0.035183, -1.044283, -2.744244, -0.923862, 1.570796, 1.605979],accel_mss,speed_ms,0,blend_radius_m)
  movel([0.032632, -1.044370, -2.744216, -0.923804, 1.570796, 1.603429],accel_mss,speed_ms,0,blend_radius_m)
  movel([0.030229, -1.044128, -2.744294, -0.923967, 1.570796, 1.601025],accel_mss,speed_ms,0,blend_radius_m)
  movel([0.027965, -1.043586, -2.744470, -0.924333, 1.570796, 1.598761],accel_mss,speed_ms,0,blend_radius_m)
  movel([0.025843, -1.042774, -2.744733, -0.924882, 1.570796, 1.596639],accel_mss,speed_ms,0,blend_radius_m)
  movel([0.023853, -1.041729, -2.745071, -0.925590, 1.570796, 1.594650],accel_mss,speed_ms,0,blend_radius_m)
  movel([0.021991, -1.040481, -2.745473, -0.926435, 1.570796, 1.592787],accel_mss,speed_ms,0,blend_radius_m)
  movel([0.020254, -1.039054, -2.745931, -0.927404, 1.570796, 1.591051],accel_mss,speed_ms,0,blend_radius_m)
  movel([0.017143, -1.035811, -2.746966, -0.929612, 1.570796, 1.587940],accel_mss,speed_ms,0,blend_radius_m)
  movel([0.014492, -1.032245, -2.748094, -0.932049, 1.570796, 1.585288],accel_mss,speed_ms,0,blend_radius_m)
  movel([0.012279, -1.028615, -2.749233, -0.934541, 1.570796, 1.583076],accel_mss,speed_ms,0,blend_radius_m)
  movel([0.010780, -1.025665, -2.750150, -0.936574, 1.570796, 1.581576],accel_mss,speed_ms,0,blend_radius_m)
  movel([0.009435, -1.022452, -2.751141, -0.938796, 1.570796, 1.580232],accel_mss,speed_ms,0,blend_radius_m)
  movel([0.008265, -1.018984, -2.752202, -0.941203, 1.570796, 1.579062],accel_mss,speed_ms,0,blend_radius_m)
  movel([0.007306, -1.015274, -2.753327, -0.943788, 1.570796, 1.578102],accel_mss,speed_ms,0,blend_radius_m)
  movel([0.006575, -1.011337, -2.754509, -0.946544, 1.570796, 1.577371],accel_mss,speed_ms,0,blend_radius_m)
  movel([0.006105, -1.007182, -2.755743, -0.949464, 1.570796, 1.576901],accel_mss,speed_ms,0,blend_radius_m)
  movel([0.005928, -1.002820, -2.757025, -0.952544, 1.570796, 1.576724],accel_mss,speed_ms,0,blend_radius_m)
  movel([0.006071, -0.998263, -2.758349, -0.955778, 1.570796, 1.576868],accel_mss,speed_ms,0,blend_radius_m)
  movel([0.006563, -0.993518, -2.759710, -0.959160, 1.570796, 1.577359],accel_mss,speed_ms,0,blend_radius_m)
  movel([0.007436, -0.988607, -2.761103, -0.962680, 1.570796, 1.578232],accel_mss,speed_ms,0,blend_radius_m)
  movel([0.008720, -0.983530, -2.762523, -0.966336, 1.570796, 1.579516],accel_mss,speed_ms,0,blend_radius_m)
  movel([0.010453, -0.978302, -2.763966, -0.970120, 1.570796, 1.581249],accel_mss,speed_ms,0,blend_radius_m)
  movel([0.012661, -0.972941, -2.765426, -0.974022, 1.570796, 1.583458],accel_mss,speed_ms,0,blend_radius_m)
  movel([0.015384, -0.967451, -2.766900, -0.978039, 1.570796, 1.586181],accel_mss,speed_ms,0,blend_radius_m)
  movel([0.018649, -0.961857, -2.768379, -0.982152, 1.570796, 1.589446],accel_mss,speed_ms,0,blend_radius_m)
  movel([0.022491, -0.956172, -2.769861, -0.986356, 1.570796, 1.593287],accel_mss,speed_ms,0,blend_radius_m)
  movel([0.024161, -0.954031, -2.770413, -0.987945, 1.570796, 1.594957],accel_mss,speed_ms,0,blend_radius_m)
  movel([0.025079, -0.953067, -2.770661, -0.988661, 1.570796, 1.595875],accel_mss,speed_ms,0,blend_radius_m)
  movel([0.026054, -0.952258, -2.770868, -0.989263, 1.570796, 1.596851],accel_mss,speed_ms,0,blend_radius_m)
  movel([0.027520, -0.951506, -2.771060, -0.989823, 1.570796, 1.598316],accel_mss,speed_ms,0,blend_radius_m)
  movel([0.028823, -0.951329, -2.771106, -0.989955, 1.570796, 1.599619],accel_mss,speed_ms,0,blend_radius_m)
  movel([0.029911, -0.951628, -2.771029, -0.989732, 1.570796, 1.600707],accel_mss,speed_ms,0,blend_radius_m)
  movel([0.030731, -0.952300, -2.770857, -0.989232, 1.570796, 1.601527],accel_mss,speed_ms,0,blend_radius_m)
  movel([0.031881, -0.954472, -2.770300, -0.987617, 1.570796, 1.602677],accel_mss,speed_ms,0,blend_radius_m)
  movel([0.032501, -0.957162, -2.769604, -0.985622, 1.570796, 1.603297],accel_mss,speed_ms,0,blend_radius_m)
  movel([0.033157, -0.962960, -2.768089, -0.981340, 1.570796, 1.603954],accel_mss,speed_ms,0,blend_radius_m)
  movel([0.033560, -0.963857, -2.767853, -0.980679, 1.570796, 1.604356],accel_mss,speed_ms,0,blend_radius_m)
  movel([0.034009, -0.963893, -2.767843, -0.980653, 1.570796, 1.604805],accel_mss,speed_ms,0,blend_radius_m)
  movel([0.034702, -0.963566, -2.767930, -0.980893, 1.570796, 1.605499],accel_mss,speed_ms,0,blend_radius_m)
  movel([0.035843, -0.960830, -2.768649, -0.982910, 1.570796, 1.606639],accel_mss,speed_ms,0,blend_radius_m)
  movel([0.036834, -0.958066, -2.769370, -0.984953, 1.570796, 1.607630],accel_mss,speed_ms,0,blend_radius_m)
  movel([0.037444, -0.966758, -2.767084, -0.978547, 1.570796, 1.608241],accel_mss,speed_ms,0,blend_radius_m)
  movel([0.038358, -0.975148, -2.764828, -0.972414, 1.570796, 1.609155],accel_mss,speed_ms,0,blend_radius_m)
  movel([0.039568, -0.983236, -2.762605, -0.966549, 1.570796, 1.610365],accel_mss,speed_ms,0,blend_radius_m)
  movel([0.041067, -0.991032, -2.760418, -0.960940, 1.570796, 1.611863],accel_mss,speed_ms,0,blend_radius_m)
  movel([0.041844, -0.994312, -2.759484, -0.958594, 1.570796, 1.612640],accel_mss,speed_ms,0,blend_radius_m)
  movel([0.042968, -0.997481, -2.758574, -0.956334, 1.570796, 1.613764],accel_mss,speed_ms,0,blend_radius_m)
  movel([0.043724, -0.998883, -2.758169, -0.955337, 1.570796, 1.614520],accel_mss,speed_ms,0,blend_radius_m)
  movel([0.044642, -1.000086, -2.757821, -0.954482, 1.570796, 1.615439],accel_mss,speed_ms,0,blend_radius_m)
  movel([0.045753, -1.001031, -2.757546, -0.953812, 1.570796, 1.616549],accel_mss,speed_ms,0,blend_radius_m)
  movel([0.047082, -1.001659, -2.757364, -0.953366, 1.570796, 1.617878],accel_mss,speed_ms,0,blend_radius_m)
  movel([0.048145, -1.001865, -2.757303, -0.953220, 1.570796, 1.618941],accel_mss,speed_ms,0,blend_radius_m)
  movel([0.050510, -1.001643, -2.757368, -0.953378, 1.570796, 1.621306],accel_mss,speed_ms,0,blend_radius_m)
  movel([0.051789, -1.001245, -2.757484, -0.953660, 1.570796, 1.622585],accel_mss,speed_ms,0,blend_radius_m)
  movel([0.054481, -0.999969, -2.757855, -0.954565, 1.570796, 1.625277],accel_mss,speed_ms,0,blend_radius_m)
  movel([0.057280, -0.998146, -2.758382, -0.955861, 1.570796, 1.628077],accel_mss,speed_ms,0,blend_radius_m)
  movel([0.060093, -0.995913, -2.759025, -0.957450, 1.570796, 1.630889],accel_mss,speed_ms,0,blend_radius_m)
  movel([0.062827, -0.993392, -2.759746, -0.959250, 1.570796, 1.633623],accel_mss,speed_ms,0,blend_radius_m)
  movel([0.065387, -0.990720, -2.760506, -0.961163, 1.570796, 1.636184],accel_mss,speed_ms,0,blend_radius_m)
  movel([0.067670, -0.988027, -2.761266, -0.963096, 1.570796, 1.638466],accel_mss,speed_ms,0,blend_radius_m)
  speed_ms = 0.005
  movel([0.067670, -0.978167, -2.755542, -0.978680, 1.570796, 1.638466],accel_mss,speed_ms,0,blend_radius_m)
  speed_ms = 0.040
  movel([0.054777, -0.986408, -2.753224, -0.972757, 1.570796, 1.625574],accel_mss,speed_ms,0,blend_radius_m)
  speed_ms = 0.005
  movel([0.054777, -0.996296, -2.758915, -0.957178, 1.570796, 1.625574],accel_mss,speed_ms,0,blend_radius_m)
  speed_ms = 0.025
  movel([0.056594, -0.994051, -2.759558, -0.958780, 1.570796, 1.627391],accel_mss,speed_ms,0,blend_radius_m)
  movel([0.060089, -0.989107, -2.760962, -0.962321, 1.570796, 1.630885],accel_mss,speed_ms,0,blend_radius_m)
  movel([0.061733, -0.986460, -2.761706, -0.964224, 1.570796, 1.632530],accel_mss,speed_ms,0,blend_radius_m)
  movel([0.064740, -0.980951, -2.763237, -0.968200, 1.570796, 1.635536],accel_mss,speed_ms,0,blend_radius_m)
  movel([0.067277, -0.975327, -2.764779, -0.972283, 1.570796, 1.638073],accel_mss,speed_ms,0,blend_radius_m)
  movel([0.068328, -0.972546, -2.765533, -0.974310, 1.570796, 1.639124],accel_mss,speed_ms,0,blend_radius_m)
  movel([0.069210, -0.969817, -2.766267, -0.976305, 1.570796, 1.640006],accel_mss,speed_ms,0,blend_radius_m)
  movel([0.070403, -0.964650, -2.767643, -0.980095, 1.570796, 1.641199],accel_mss,speed_ms,0,blend_radius_m)
  movel([0.070684, -0.962266, -2.768272, -0.981851, 1.570796, 1.641480],accel_mss,speed_ms,0,blend_radius_m)
  movel([0.070726, -0.960063, -2.768849, -0.983477, 1.570796, 1.641522],accel_mss,speed_ms,0,blend_radius_m)
  movel([0.070518, -0.958066, -2.769370, -0.984953, 1.570796, 1.641314],accel_mss,speed_ms,0,blend_radius_m)
  movel([0.070039, -0.956305, -2.769826, -0.986257, 1.570796, 1.640836],accel_mss,speed_ms,0,blend_radius_m)
  movel([0.069145, -0.954396, -2.770319, -0.987674, 1.570796, 1.639941],accel_mss,speed_ms,0,blend_radius_m)
  movel([0.067993, -0.952760, -2.770739, -0.988889, 1.570796, 1.638790],accel_mss,speed_ms,0,blend_radius_m)
  movel([0.066567, -0.951475, -2.771068, -0.989845, 1.570796, 1.637363],accel_mss,speed_ms,0,blend_radius_m)
  movel([0.064853, -0.950624, -2.771285, -0.990479, 1.570796, 1.635649],accel_mss,speed_ms,0,blend_radius_m)
  movel([0.062833, -0.950283, -2.771372, -0.990733, 1.570796, 1.633630],accel_mss,speed_ms,0,blend_radius_m)
  movel([0.060502, -0.950531, -2.771309, -0.990549, 1.570796, 1.631299],accel_mss,speed_ms,0,blend_radius_m)
  movel([0.057846, -0.951444, -2.771076, -0.989869, 1.570796, 1.628642],accel_mss,speed_ms,0,blend_radius_m)
  movel([0.054857, -0.953088, -2.770655, -0.988646, 1.570796, 1.625654],accel_mss,speed_ms,0,blend_radius_m)
  movel([0.052795, -0.954596, -2.770268, -0.987525, 1.570796, 1.623592],accel_mss,speed_ms,0,blend_radius_m)
  movel([0.050789, -0.956398, -2.769802, -0.986189, 1.570796, 1.621585],accel_mss,speed_ms,0,blend_radius_m)
  movel([0.048907, -0.958416, -2.769279, -0.984694, 1.570796, 1.619703],accel_mss,speed_ms,0,blend_radius_m)
  movel([0.047206, -0.960580, -2.768714, -0.983095, 1.570796, 1.618002],accel_mss,speed_ms,0,blend_radius_m)
  movel([0.045744, -0.962820, -2.768126, -0.981443, 1.570796, 1.616540],accel_mss,speed_ms,0,blend_radius_m)
  movel([0.044580, -0.965064, -2.767534, -0.979791, 1.570796, 1.615376],accel_mss,speed_ms,0,blend_radius_m)
  movel([0.043774, -0.967243, -2.766955, -0.978191, 1.570796, 1.614571],accel_mss,speed_ms,0,blend_radius_m)
  movel([0.043376, -0.969292, -2.766408, -0.976689, 1.570796, 1.614172],accel_mss,speed_ms,0,blend_radius_m)
  speed_ms = 0.005
  movel([0.043376, -0.959505, -2.760610, -0.992274, 1.570796, 1.614172],accel_mss,speed_ms,0,blend_radius_m)
  speed_ms = 0.040
  # Splitting Linear movement in 2 (instruction 399: MoveL 378)
  movel([0.095251, -0.966227, -2.758813, -0.987349, 1.570796, 1.666048],accel_mss,speed_ms,0,blend_radius_m)
  movel([0.144369, -0.976923, -2.755887, -0.979579, 1.570796, 1.715166],accel_mss,speed_ms,0,blend_radius_m)
  speed_ms = 0.005
  movel([0.144369, -0.986778, -2.761616, -0.963994, 1.570796, 1.715166],accel_mss,speed_ms,0,blend_radius_m)
  speed_ms = 0.025
  movel([0.142576, -0.997367, -2.758607, -0.956415, 1.570796, 1.713373],accel_mss,speed_ms,0,blend_radius_m)
  movel([0.141323, -1.002736, -2.757049, -0.952604, 1.570796, 1.712119],accel_mss,speed_ms,0,blend_radius_m)
  movel([0.140478, -1.005508, -2.756237, -0.950645, 1.570796, 1.711274],accel_mss,speed_ms,0,blend_radius_m)
  movel([0.139439, -1.008358, -2.755395, -0.948636, 1.570796, 1.710235],accel_mss,speed_ms,0,blend_radius_m)
  movel([0.138085, -1.011421, -2.754483, -0.946484, 1.570796, 1.708881],accel_mss,speed_ms,0,blend_radius_m)
  movel([0.137248, -1.012938, -2.754029, -0.945421, 1.570796, 1.708044],accel_mss,speed_ms,0,blend_radius_m)
  movel([0.136253, -1.014420, -2.753584, -0.944385, 1.570796, 1.707050],accel_mss,speed_ms,0,blend_radius_m)
  movel([0.136298, -1.012112, -2.754277, -0.946000, 1.570796, 1.707094],accel_mss,speed_ms,0,blend_radius_m)
  movel([0.135952, -1.010059, -2.754890, -0.947440, 1.570796, 1.706749],accel_mss,speed_ms,0,blend_radius_m)
  movel([0.135606, -1.009554, -2.755040, -0.947795, 1.570796, 1.706403],accel_mss,speed_ms,0,blend_radius_m)
  movel([0.135231, -1.009599, -2.755027, -0.947763, 1.570796, 1.706027],accel_mss,speed_ms,0,blend_radius_m)
  movel([0.134795, -1.009848, -2.754953, -0.947589, 1.570796, 1.705592],accel_mss,speed_ms,0,blend_radius_m)
  movel([0.133917, -1.010689, -2.754702, -0.946998, 1.570796, 1.704713],accel_mss,speed_ms,0,blend_radius_m)
  movel([0.132686, -1.012289, -2.754224, -0.945876, 1.570796, 1.703482],accel_mss,speed_ms,0,blend_radius_m)
  movel([0.131708, -1.013891, -2.753743, -0.944755, 1.570796, 1.702505],accel_mss,speed_ms,0,blend_radius_m)
  movel([0.130937, -1.015487, -2.753262, -0.943639, 1.570796, 1.701733],accel_mss,speed_ms,0,blend_radius_m)
  movel([0.130326, -1.017073, -2.752783, -0.942533, 1.570796, 1.701122],accel_mss,speed_ms,0,blend_radius_m)
  movel([0.128511, -1.023321, -2.750874, -0.938194, 1.570796, 1.699307],accel_mss,speed_ms,0,blend_radius_m)
  movel([0.127266, -1.027012, -2.749732, -0.935645, 1.570796, 1.698062],accel_mss,speed_ms,0,blend_radius_m)
  movel([0.125795, -1.030729, -2.748571, -0.933089, 1.570796, 1.696591],accel_mss,speed_ms,0,blend_radius_m)
  movel([0.124038, -1.034457, -2.747396, -0.930537, 1.570796, 1.694835],accel_mss,speed_ms,0,blend_radius_m)
  movel([0.121941, -1.038161, -2.746217, -0.928011, 1.570796, 1.692737],accel_mss,speed_ms,0,blend_radius_m)
  movel([0.122563, -1.035397, -2.747098, -0.929894, 1.570796, 1.693359],accel_mss,speed_ms,0,blend_radius_m)
  movel([0.122553, -1.032931, -2.747878, -0.931580, 1.570796, 1.693350],accel_mss,speed_ms,0,blend_radius_m)
  movel([0.122409, -1.032399, -2.748046, -0.931944, 1.570796, 1.693205],accel_mss,speed_ms,0,blend_radius_m)
  movel([0.122040, -1.032106, -2.748138, -0.932145, 1.570796, 1.692837],accel_mss,speed_ms,0,blend_radius_m)
  movel([0.121554, -1.032190, -2.748112, -0.932087, 1.570796, 1.692350],accel_mss,speed_ms,0,blend_radius_m)
  movel([0.121001, -1.032524, -2.748007, -0.931859, 1.570796, 1.691797],accel_mss,speed_ms,0,blend_radius_m)
  movel([0.119921, -1.033581, -2.747673, -0.931135, 1.570796, 1.690717],accel_mss,speed_ms,0,blend_radius_m)
  movel([0.118765, -1.035100, -2.747192, -0.930097, 1.570796, 1.689561],accel_mss,speed_ms,0,blend_radius_m)
  movel([0.117777, -1.036679, -2.746690, -0.929020, 1.570796, 1.688573],accel_mss,speed_ms,0,blend_radius_m)
  movel([0.116176, -1.039924, -2.745652, -0.926813, 1.570796, 1.686972],accel_mss,speed_ms,0,blend_radius_m)
  movel([0.113543, -1.046316, -2.743582, -0.922491, 1.570796, 1.684339],accel_mss,speed_ms,0,blend_radius_m)
  movel([0.111823, -1.049874, -2.742415, -0.920099, 1.570796, 1.682619],accel_mss,speed_ms,0,blend_radius_m)
  movel([0.109889, -1.053410, -2.741246, -0.917733, 1.570796, 1.680686],accel_mss,speed_ms,0,blend_radius_m)
  movel([0.107694, -1.056874, -2.740090, -0.915425, 1.570796, 1.678490],accel_mss,speed_ms,0,blend_radius_m)
  movel([0.105191, -1.060220, -2.738964, -0.913205, 1.570796, 1.675988],accel_mss,speed_ms,0,blend_radius_m)
  movel([0.105698, -1.058700, -2.739477, -0.914213, 1.570796, 1.676494],accel_mss,speed_ms,0,blend_radius_m)
  movel([0.106188, -1.055838, -2.740437, -0.916114, 1.570796, 1.676984],accel_mss,speed_ms,0,blend_radius_m)
  movel([0.106161, -1.054539, -2.740870, -0.916980, 1.570796, 1.676958],accel_mss,speed_ms,0,blend_radius_m)
  movel([0.106006, -1.054029, -2.741040, -0.917320, 1.570796, 1.676802],accel_mss,speed_ms,0,blend_radius_m)
  movel([0.105552, -1.053924, -2.741075, -0.917390, 1.570796, 1.676348],accel_mss,speed_ms,0,blend_radius_m)
  movel([0.104890, -1.054438, -2.740904, -0.917047, 1.570796, 1.675687],accel_mss,speed_ms,0,blend_radius_m)
  movel([0.103405, -1.056078, -2.740357, -0.915955, 1.570796, 1.674202],accel_mss,speed_ms,0,blend_radius_m)
  movel([0.102119, -1.057745, -2.739798, -0.914846, 1.570796, 1.672915],accel_mss,speed_ms,0,blend_radius_m)
  movel([0.099909, -1.061147, -2.738650, -0.912592, 1.570796, 1.670705],accel_mss,speed_ms,0,blend_radius_m)
  movel([0.097790, -1.064577, -2.737483, -0.910329, 1.570796, 1.668586],accel_mss,speed_ms,0,blend_radius_m)
  movel([0.096618, -1.066288, -2.736897, -0.909204, 1.570796, 1.667414],accel_mss,speed_ms,0,blend_radius_m)
  movel([0.095292, -1.067988, -2.736313, -0.908088, 1.570796, 1.666088],accel_mss,speed_ms,0,blend_radius_m)
  movel([0.091838, -1.071925, -2.734950, -0.905515, 1.570796, 1.662635],accel_mss,speed_ms,0,blend_radius_m)
  movel([0.088265, -1.075713, -2.733625, -0.903051, 1.570796, 1.659061],accel_mss,speed_ms,0,blend_radius_m)
  movel([0.084609, -1.079357, -2.732340, -0.900692, 1.570796, 1.655405],accel_mss,speed_ms,0,blend_radius_m)
  movel([0.080897, -1.082880, -2.731085, -0.898423, 1.570796, 1.651693],accel_mss,speed_ms,0,blend_radius_m)
  speed_ms = 0.005
  movel([0.080897, -1.072849, -2.725755, -0.913784, 1.570796, 1.651693],accel_mss,speed_ms,0,blend_radius_m)
  speed_ms = 0.040
  movel([0.052585, -1.044492, -2.735430, -0.932467, 1.570796, 1.623381],accel_mss,speed_ms,0,blend_radius_m)
  speed_ms = 0.005
  movel([0.052585, -1.054505, -2.740881, -0.917002, 1.570796, 1.623381],accel_mss,speed_ms,0,blend_radius_m)
  speed_ms = 0.025
  movel([0.053739, -1.053150, -2.741332, -0.917907, 1.570796, 1.624535],accel_mss,speed_ms,0,blend_radius_m)
  movel([0.054770, -1.051675, -2.741821, -0.918893, 1.570796, 1.625566],accel_mss,speed_ms,0,blend_radius_m)
  movel([0.056627, -1.048500, -2.742867, -0.921022, 1.570796, 1.627423],accel_mss,speed_ms,0,blend_radius_m)
  movel([0.058462, -1.045248, -2.743930, -0.923211, 1.570796, 1.629259],accel_mss,speed_ms,0,blend_radius_m)
  movel([0.059472, -1.043675, -2.744441, -0.924273, 1.570796, 1.630269],accel_mss,speed_ms,0,blend_radius_m)
  movel([0.060595, -1.042184, -2.744924, -0.925281, 1.570796, 1.631391],accel_mss,speed_ms,0,blend_radius_m)
  movel([0.061493, -1.041195, -2.745243, -0.925951, 1.570796, 1.632289],accel_mss,speed_ms,0,blend_radius_m)
  movel([0.062238, -1.040561, -2.745447, -0.926381, 1.570796, 1.633034],accel_mss,speed_ms,0,blend_radius_m)
  movel([0.062844, -1.040241, -2.745550, -0.926598, 1.570796, 1.633640],accel_mss,speed_ms,0,blend_radius_m)
  movel([0.063327, -1.040198, -2.745564, -0.926627, 1.570796, 1.634123],accel_mss,speed_ms,0,blend_radius_m)
  movel([0.063959, -1.040814, -2.745366, -0.926209, 1.570796, 1.634756],accel_mss,speed_ms,0,blend_radius_m)
  movel([0.064238, -1.042108, -2.744948, -0.925332, 1.570796, 1.635035],accel_mss,speed_ms,0,blend_radius_m)
  movel([0.064127, -1.045569, -2.743826, -0.922994, 1.570796, 1.634924],accel_mss,speed_ms,0,blend_radius_m)
  movel([0.063808, -1.048251, -2.742949, -0.921189, 1.570796, 1.634605],accel_mss,speed_ms,0,blend_radius_m)
  movel([0.065855, -1.045006, -2.744009, -0.923374, 1.570796, 1.636651],accel_mss,speed_ms,0,blend_radius_m)
  movel([0.067407, -1.041899, -2.745016, -0.925474, 1.570796, 1.638203],accel_mss,speed_ms,0,blend_radius_m)
  movel([0.068592, -1.038883, -2.745986, -0.927520, 1.570796, 1.639389],accel_mss,speed_ms,0,blend_radius_m)
  movel([0.069527, -1.035924, -2.746930, -0.929535, 1.570796, 1.640323],accel_mss,speed_ms,0,blend_radius_m)
  movel([0.072078, -1.026949, -2.749752, -0.935688, 1.570796, 1.642875],accel_mss,speed_ms,0,blend_radius_m)
  movel([0.073262, -1.023779, -2.750733, -0.937877, 1.570796, 1.644059],accel_mss,speed_ms,0,blend_radius_m)
  movel([0.073925, -1.022484, -2.751131, -0.938773, 1.570796, 1.644722],accel_mss,speed_ms,0,blend_radius_m)
  movel([0.074609, -1.021646, -2.751389, -0.939354, 1.570796, 1.645405],accel_mss,speed_ms,0,blend_radius_m)
  movel([0.075288, -1.021199, -2.751526, -0.939664, 1.570796, 1.646084],accel_mss,speed_ms,0,blend_radius_m)
  movel([0.075933, -1.021087, -2.751560, -0.939742, 1.570796, 1.646729],accel_mss,speed_ms,0,blend_radius_m)
  movel([0.076523, -1.021240, -2.751513, -0.939635, 1.570796, 1.647320],accel_mss,speed_ms,0,blend_radius_m)
  movel([0.077028, -1.021600, -2.751403, -0.939386, 1.570796, 1.647824],accel_mss,speed_ms,0,blend_radius_m)
  movel([0.077688, -1.022679, -2.751071, -0.938638, 1.570796, 1.648484],accel_mss,speed_ms,0,blend_radius_m)
  movel([0.077828, -1.024123, -2.750627, -0.937639, 1.570796, 1.648624],accel_mss,speed_ms,0,blend_radius_m)
  movel([0.077674, -1.026131, -2.750005, -0.936252, 1.570796, 1.648471],accel_mss,speed_ms,0,blend_radius_m)
  movel([0.077147, -1.029933, -2.748821, -0.933636, 1.570796, 1.647943],accel_mss,speed_ms,0,blend_radius_m)
  movel([0.079247, -1.023727, -2.750749, -0.937913, 1.570796, 1.650044],accel_mss,speed_ms,0,blend_radius_m)
  movel([0.080045, -1.020682, -2.751684, -0.940023, 1.570796, 1.650842],accel_mss,speed_ms,0,blend_radius_m)
  movel([0.081117, -1.014760, -2.753482, -0.944147, 1.570796, 1.651913],accel_mss,speed_ms,0,blend_radius_m)
  movel([0.081382, -1.011915, -2.754336, -0.946138, 1.570796, 1.652178],accel_mss,speed_ms,0,blend_radius_m)
  movel([0.081355, -1.006515, -2.755940, -0.949934, 1.570796, 1.652151],accel_mss,speed_ms,0,blend_radius_m)
  speed_ms = 0.005
  movel([0.081355, -0.996596, -2.750290, -0.965503, 1.570796, 1.652151],accel_mss,speed_ms,0,blend_radius_m)
  speed_ms = 0.040
  movel([0.062258, -1.022904, -2.742351, -0.947135, 1.570796, 1.633054],accel_mss,speed_ms,0,blend_radius_m)
  speed_ms = 0.005
  movel([0.062258, -1.032885, -2.747893, -0.931611, 1.570796, 1.633054],accel_mss,speed_ms,0,blend_radius_m)
  speed_ms = 0.025
  movel([0.059858, -1.036607, -2.746713, -0.929069, 1.570796, 1.630654],accel_mss,speed_ms,0,blend_radius_m)
  movel([0.057669, -1.040351, -2.745514, -0.926523, 1.570796, 1.628466],accel_mss,speed_ms,0,blend_radius_m)
  movel([0.053440, -1.047798, -2.743097, -0.921493, 1.570796, 1.624237],accel_mss,speed_ms,0,blend_radius_m)
  movel([0.051127, -1.051479, -2.741886, -0.919024, 1.570796, 1.621923],accel_mss,speed_ms,0,blend_radius_m)
  movel([0.048566, -1.055047, -2.740701, -0.916641, 1.570796, 1.619362],accel_mss,speed_ms,0,blend_radius_m)
  movel([0.045728, -1.058361, -2.739591, -0.914437, 1.570796, 1.616525],accel_mss,speed_ms,0,blend_radius_m)
  movel([0.044200, -1.059878, -2.739079, -0.913431, 1.570796, 1.614997],accel_mss,speed_ms,0,blend_radius_m)
  movel([0.042596, -1.061281, -2.738605, -0.912503, 1.570796, 1.613392],accel_mss,speed_ms,0,blend_radius_m)
  movel([0.043768, -1.060024, -2.739030, -0.913335, 1.570796, 1.614565],accel_mss,speed_ms,0,blend_radius_m)
  movel([0.044992, -1.058212, -2.739641, -0.914536, 1.570796, 1.615788],accel_mss,speed_ms,0,blend_radius_m)
  movel([0.046127, -1.056100, -2.740349, -0.915940, 1.570796, 1.616923],accel_mss,speed_ms,0,blend_radius_m)
  movel([0.047012, -1.053957, -2.741064, -0.917368, 1.570796, 1.617809],accel_mss,speed_ms,0,blend_radius_m)
  movel([0.047502, -1.052041, -2.741700, -0.918648, 1.570796, 1.618298],accel_mss,speed_ms,0,blend_radius_m)
  movel([0.047545, -1.051260, -2.741958, -0.919171, 1.570796, 1.618341],accel_mss,speed_ms,0,blend_radius_m)
  movel([0.047433, -1.050636, -2.742165, -0.919589, 1.570796, 1.618230],accel_mss,speed_ms,0,blend_radius_m)
  movel([0.047146, -1.050202, -2.742307, -0.919879, 1.570796, 1.617942],accel_mss,speed_ms,0,blend_radius_m)
  movel([0.046658, -1.050000, -2.742374, -0.920015, 1.570796, 1.617455],accel_mss,speed_ms,0,blend_radius_m)
  movel([0.045960, -1.050056, -2.742356, -0.919977, 1.570796, 1.616756],accel_mss,speed_ms,0,blend_radius_m)
  movel([0.045023, -1.050409, -2.742239, -0.919741, 1.570796, 1.615819],accel_mss,speed_ms,0,blend_radius_m)
  movel([0.043517, -1.051438, -2.741899, -0.919051, 1.570796, 1.614313],accel_mss,speed_ms,0,blend_radius_m)
  movel([0.037327, -1.057006, -2.740046, -0.915337, 1.570796, 1.608124],accel_mss,speed_ms,0,blend_radius_m)
  movel([0.034681, -1.059116, -2.739336, -0.913937, 1.570796, 1.605478],accel_mss,speed_ms,0,blend_radius_m)
  movel([0.031966, -1.061059, -2.738680, -0.912650, 1.570796, 1.602762],accel_mss,speed_ms,0,blend_radius_m)
  movel([0.029266, -1.062729, -2.738113, -0.911547, 1.570796, 1.600063],accel_mss,speed_ms,0,blend_radius_m)
  movel([0.026666, -1.064006, -2.737678, -0.910705, 1.570796, 1.597462],accel_mss,speed_ms,0,blend_radius_m)
  movel([0.024244, -1.064783, -2.737413, -0.910193, 1.570796, 1.595040],accel_mss,speed_ms,0,blend_radius_m)
  movel([0.022086, -1.064937, -2.737360, -0.910092, 1.570796, 1.592882],accel_mss,speed_ms,0,blend_radius_m)
  movel([0.022777, -1.064780, -2.737414, -0.910195, 1.570796, 1.593573],accel_mss,speed_ms,0,blend_radius_m)
  movel([0.023686, -1.064263, -2.737590, -0.910535, 1.570796, 1.594482],accel_mss,speed_ms,0,blend_radius_m)
  movel([0.025867, -1.062522, -2.738183, -0.911683, 1.570796, 1.596664],accel_mss,speed_ms,0,blend_radius_m)
  movel([0.028010, -1.060454, -2.738885, -0.913051, 1.570796, 1.598806],accel_mss,speed_ms,0,blend_radius_m)
  movel([0.029486, -1.058809, -2.739440, -0.914140, 1.570796, 1.600282],accel_mss,speed_ms,0,blend_radius_m)
  movel([0.030353, -1.057552, -2.739862, -0.914974, 1.570796, 1.601149],accel_mss,speed_ms,0,blend_radius_m)
  movel([0.030677, -1.056722, -2.740141, -0.915526, 1.570796, 1.601473],accel_mss,speed_ms,0,blend_radius_m)
  movel([0.030544, -1.056251, -2.740299, -0.915839, 1.570796, 1.601341],accel_mss,speed_ms,0,blend_radius_m)
  movel([0.030055, -1.056072, -2.740358, -0.915958, 1.570796, 1.600851],accel_mss,speed_ms,0,blend_radius_m)
  movel([0.028394, -1.056321, -2.740275, -0.915793, 1.570796, 1.599190],accel_mss,speed_ms,0,blend_radius_m)
  movel([0.026468, -1.056924, -2.740073, -0.915392, 1.570796, 1.597264],accel_mss,speed_ms,0,blend_radius_m)
  movel([0.022092, -1.058291, -2.739614, -0.914484, 1.570796, 1.592888],accel_mss,speed_ms,0,blend_radius_m)
  movel([0.017739, -1.059280, -2.739281, -0.913828, 1.570796, 1.588535],accel_mss,speed_ms,0,blend_radius_m)
  movel([0.015686, -1.059498, -2.739208, -0.913683, 1.570796, 1.586482],accel_mss,speed_ms,0,blend_radius_m)
  movel([0.013777, -1.059457, -2.739221, -0.913710, 1.570796, 1.584574],accel_mss,speed_ms,0,blend_radius_m)
  movel([0.012060, -1.059101, -2.739342, -0.913947, 1.570796, 1.582856],accel_mss,speed_ms,0,blend_radius_m)
  movel([0.010581, -1.058374, -2.739586, -0.914429, 1.570796, 1.581377],accel_mss,speed_ms,0,blend_radius_m)
  movel([0.013190, -1.057531, -2.739870, -0.914989, 1.570796, 1.583987],accel_mss,speed_ms,0,blend_radius_m)
  movel([0.014621, -1.056760, -2.740128, -0.915501, 1.570796, 1.585417],accel_mss,speed_ms,0,blend_radius_m)
  movel([0.015257, -1.056256, -2.740297, -0.915836, 1.570796, 1.586053],accel_mss,speed_ms,0,blend_radius_m)
  movel([0.015800, -1.055655, -2.740498, -0.916236, 1.570796, 1.586596],accel_mss,speed_ms,0,blend_radius_m)
  movel([0.016023, -1.055197, -2.740651, -0.916541, 1.570796, 1.586820],accel_mss,speed_ms,0,blend_radius_m)
  movel([0.015994, -1.054782, -2.740789, -0.916818, 1.570796, 1.586790],accel_mss,speed_ms,0,blend_radius_m)
  movel([0.015315, -1.054072, -2.741026, -0.917291, 1.570796, 1.586112],accel_mss,speed_ms,0,blend_radius_m)
  movel([0.013996, -1.053512, -2.741212, -0.917665, 1.570796, 1.584792],accel_mss,speed_ms,0,blend_radius_m)
  movel([0.012280, -1.053078, -2.741356, -0.917955, 1.570796, 1.583076],accel_mss,speed_ms,0,blend_radius_m)
  movel([0.006259, -1.052217, -2.741642, -0.918530, 1.570796, 1.577055],accel_mss,speed_ms,0,blend_radius_m)
  movel([0.004079, -1.051553, -2.741862, -0.918975, 1.570796, 1.574875],accel_mss,speed_ms,0,blend_radius_m)
  movel([0.002111, -1.050582, -2.742182, -0.919625, 1.570796, 1.572908],accel_mss,speed_ms,0,blend_radius_m)
  movel([0.000486, -1.049216, -2.742632, -0.920541, 1.570796, 1.571283],accel_mss,speed_ms,0,blend_radius_m)
  movel([-0.000685, -1.047374, -2.743236, -0.921778, 1.570796, 1.570112],accel_mss,speed_ms,0,blend_radius_m)
  movel([0.001330, -1.048109, -2.742995, -0.921284, 1.570796, 1.572126],accel_mss,speed_ms,0,blend_radius_m)
  movel([0.002588, -1.048232, -2.742955, -0.921202, 1.570796, 1.573385],accel_mss,speed_ms,0,blend_radius_m)
  movel([0.003813, -1.047916, -2.743059, -0.921414, 1.570796, 1.574610],accel_mss,speed_ms,0,blend_radius_m)
  movel([0.004986, -1.047085, -2.743331, -0.921973, 1.570796, 1.575782],accel_mss,speed_ms,0,blend_radius_m)
  movel([0.005693, -1.046112, -2.743649, -0.922629, 1.570796, 1.576489],accel_mss,speed_ms,0,blend_radius_m)
  movel([0.005907, -1.045127, -2.743970, -0.923292, 1.570796, 1.576703],accel_mss,speed_ms,0,blend_radius_m)
  movel([0.005604, -1.044257, -2.744252, -0.923880, 1.570796, 1.576400],accel_mss,speed_ms,0,blend_radius_m)
  movel([0.003068, -1.040321, -2.745524, -0.926543, 1.570796, 1.573864],accel_mss,speed_ms,0,blend_radius_m)
  movel([0.001141, -1.035957, -2.746920, -0.929513, 1.570796, 1.571937],accel_mss,speed_ms,0,blend_radius_m)
  movel([0.000453, -1.033540, -2.747686, -0.931163, 1.570796, 1.571250],accel_mss,speed_ms,0,blend_radius_m)
  movel([-0.000030, -1.030929, -2.748508, -0.932952, 1.570796, 1.570766],accel_mss,speed_ms,0,blend_radius_m)
  movel([-0.000289, -1.028093, -2.749396, -0.934901, 1.570796, 1.570507],accel_mss,speed_ms,0,blend_radius_m)
  movel([-0.000305, -1.025000, -2.750356, -0.937033, 1.570796, 1.570491],accel_mss,speed_ms,0,blend_radius_m)
  speed_ms = 0.005
  movel([-0.000305, -1.015035, -2.744781, -0.952573, 1.570796, 1.570491],accel_mss,speed_ms,0,blend_radius_m)
  speed_ms = 0.040
  movel([-0.041269, -1.007422, -2.747087, -0.957880, 1.570796, 1.529527],accel_mss,speed_ms,0,blend_radius_m)
  speed_ms = 0.005
  movel([-0.041269, -1.017369, -2.752693, -0.942327, 1.570796, 1.529527],accel_mss,speed_ms,0,blend_radius_m)
  speed_ms = 0.025
  movel([-0.037935, -1.011786, -2.754375, -0.946229, 1.570796, 1.532862],accel_mss,speed_ms,0,blend_radius_m)
  movel([-0.034722, -1.006144, -2.756049, -0.950196, 1.570796, 1.536074],accel_mss,speed_ms,0,blend_radius_m)
  movel([-0.028597, -0.994653, -2.759386, -0.958350, 1.570796, 1.542199],accel_mss,speed_ms,0,blend_radius_m)
  movel([-0.022885, -0.982918, -2.762693, -0.966778, 1.570796, 1.547912],accel_mss,speed_ms,0,blend_radius_m)
  movel([-0.017602, -0.970978, -2.765955, -0.975456, 1.570796, 1.553194],accel_mss,speed_ms,0,blend_radius_m)
  movel([-0.012765, -0.958869, -2.769161, -0.984359, 1.570796, 1.558032],accel_mss,speed_ms,0,blend_radius_m)
  movel([-0.008393, -0.946637, -2.772296, -0.993456, 1.570796, 1.562403],accel_mss,speed_ms,0,blend_radius_m)
  movel([-0.004507, -0.934336, -2.775348, -1.002706, 1.570796, 1.566289],accel_mss,speed_ms,0,blend_radius_m)
  movel([-0.001128, -0.922011, -2.778305, -1.012073, 1.570796, 1.569668],accel_mss,speed_ms,0,blend_radius_m)
  movel([0.001717, -0.909732, -2.781154, -1.021503, 1.570796, 1.572514],accel_mss,speed_ms,0,blend_radius_m)
  movel([0.004003, -0.897559, -2.783885, -1.030945, 1.570796, 1.574800],accel_mss,speed_ms,0,blend_radius_m)
  movel([0.005699, -0.885564, -2.786488, -1.040337, 1.570796, 1.576495],accel_mss,speed_ms,0,blend_radius_m)
  movel([0.006772, -0.873825, -2.788951, -1.049614, 1.570796, 1.577568],accel_mss,speed_ms,0,blend_radius_m)
  movel([0.007201, -0.862408, -2.791269, -1.058712, 1.570796, 1.577998],accel_mss,speed_ms,0,blend_radius_m)
  movel([0.006944, -0.851412, -2.793431, -1.067546, 1.570796, 1.577741],accel_mss,speed_ms,0,blend_radius_m)
  movel([0.005975, -0.840920, -2.795430, -1.076039, 1.570796, 1.576771],accel_mss,speed_ms,0,blend_radius_m)
  movel([0.003369, -0.826072, -2.798156, -1.088160, 1.570796, 1.574166],accel_mss,speed_ms,0,blend_radius_m)
  movel([0.003313, -0.823298, -2.798652, -1.090439, 1.570796, 1.574110],accel_mss,speed_ms,0,blend_radius_m)
  movel([0.003753, -0.820180, -2.799205, -1.093004, 1.570796, 1.574550],accel_mss,speed_ms,0,blend_radius_m)
  movel([0.005074, -0.815499, -2.800025, -1.096865, 1.570796, 1.575870],accel_mss,speed_ms,0,blend_radius_m)
  movel([0.006722, -0.811606, -2.800698, -1.100085, 1.570796, 1.577519],accel_mss,speed_ms,0,blend_radius_m)
  movel([0.007652, -0.809945, -2.800983, -1.101461, 1.570796, 1.578448],accel_mss,speed_ms,0,blend_radius_m)
  movel([0.009696, -0.807142, -2.801460, -1.103787, 1.570796, 1.580493],accel_mss,speed_ms,0,blend_radius_m)
  movel([0.010791, -0.806000, -2.801654, -1.104736, 1.570796, 1.581587],accel_mss,speed_ms,0,blend_radius_m)
  movel([0.013113, -0.804180, -2.801960, -1.106249, 1.570796, 1.583910],accel_mss,speed_ms,0,blend_radius_m)
  movel([0.015556, -0.802943, -2.802168, -1.107278, 1.570796, 1.586352],accel_mss,speed_ms,0,blend_radius_m)
  movel([0.018066, -0.802235, -2.802286, -1.107868, 1.570796, 1.588863],accel_mss,speed_ms,0,blend_radius_m)
  movel([0.020598, -0.801998, -2.802326, -1.108065, 1.570796, 1.591395],accel_mss,speed_ms,0,blend_radius_m)
  movel([0.023097, -0.802170, -2.802297, -1.107922, 1.570796, 1.593894],accel_mss,speed_ms,0,blend_radius_m)
  movel([0.025518, -0.802695, -2.802209, -1.107485, 1.570796, 1.596315],accel_mss,speed_ms,0,blend_radius_m)
  movel([0.029924, -0.804533, -2.801901, -1.105955, 1.570796, 1.600720],accel_mss,speed_ms,0,blend_radius_m)
  movel([0.033447, -0.807004, -2.801484, -1.103901, 1.570796, 1.604244],accel_mss,speed_ms,0,blend_radius_m)
  movel([0.035752, -0.809556, -2.801049, -1.101783, 1.570796, 1.606548],accel_mss,speed_ms,0,blend_radius_m)
  movel([0.037774, -0.813243, -2.800416, -1.098730, 1.570796, 1.608570],accel_mss,speed_ms,0,blend_radius_m)
  movel([0.039406, -0.817332, -2.799705, -1.095352, 1.570796, 1.610203],accel_mss,speed_ms,0,blend_radius_m)
  movel([0.041880, -0.826262, -2.798122, -1.088005, 1.570796, 1.612676],accel_mss,speed_ms,0,blend_radius_m)
  movel([0.043907, -0.835511, -2.796437, -1.080441, 1.570796, 1.614703],accel_mss,speed_ms,0,blend_radius_m)
  movel([0.046189, -0.844293, -2.794794, -1.073301, 1.570796, 1.616985],accel_mss,speed_ms,0,blend_radius_m)
  movel([0.048787, -0.851584, -2.793398, -1.067407, 1.570796, 1.619584],accel_mss,speed_ms,0,blend_radius_m)
  movel([0.050495, -0.854778, -2.792776, -1.064835, 1.570796, 1.621292],accel_mss,speed_ms,0,blend_radius_m)
  movel([0.052701, -0.857403, -2.792262, -1.062725, 1.570796, 1.623497],accel_mss,speed_ms,0,blend_radius_m)
  movel([0.054025, -0.858266, -2.792091, -1.062031, 1.570796, 1.624822],accel_mss,speed_ms,0,blend_radius_m)
  movel([0.054860, -0.858428, -2.792059, -1.061902, 1.570796, 1.625656],accel_mss,speed_ms,0,blend_radius_m)
  movel([0.055847, -0.858300, -2.792085, -1.062004, 1.570796, 1.626643],accel_mss,speed_ms,0,blend_radius_m)
  movel([0.057282, -0.857654, -2.792212, -1.062522, 1.570796, 1.628078],accel_mss,speed_ms,0,blend_radius_m)
  movel([0.058791, -0.856588, -2.792422, -1.063379, 1.570796, 1.629587],accel_mss,speed_ms,0,blend_radius_m)
  movel([0.061813, -0.853741, -2.792979, -1.065670, 1.570796, 1.632609],accel_mss,speed_ms,0,blend_radius_m)
  movel([0.065119, -0.850113, -2.793682, -1.068594, 1.570796, 1.635915],accel_mss,speed_ms,0,blend_radius_m)
  movel([0.068277, -0.846328, -2.794407, -1.071654, 1.570796, 1.639073],accel_mss,speed_ms,0,blend_radius_m)
  movel([0.074274, -0.838388, -2.795904, -1.078098, 1.570796, 1.645070],accel_mss,speed_ms,0,blend_radius_m)
  movel([0.085956, -0.821835, -2.798912, -1.091642, 1.570796, 1.656752],accel_mss,speed_ms,0,blend_radius_m)
  movel([0.091724, -0.814088, -2.800270, -1.098031, 1.570796, 1.662520],accel_mss,speed_ms,0,blend_radius_m)
  movel([0.095118, -0.809881, -2.800994, -1.101514, 1.570796, 1.665914],accel_mss,speed_ms,0,blend_radius_m)
  movel([0.098550, -0.806072, -2.801641, -1.104675, 1.570796, 1.669346],accel_mss,speed_ms,0,blend_radius_m)
  movel([0.100208, -0.804460, -2.801913, -1.106016, 1.570796, 1.671005],accel_mss,speed_ms,0,blend_radius_m)
  movel([0.101792, -0.803123, -2.802138, -1.107129, 1.570796, 1.672589],accel_mss,speed_ms,0,blend_radius_m)
  movel([0.103267, -0.802120, -2.802305, -1.107964, 1.570796, 1.674063],accel_mss,speed_ms,0,blend_radius_m)
  movel([0.104605, -0.801513, -2.802406, -1.108469, 1.570796, 1.675402],accel_mss,speed_ms,0,blend_radius_m)
  movel([0.105774, -0.801358, -2.802432, -1.108599, 1.570796, 1.676571],accel_mss,speed_ms,0,blend_radius_m)
  movel([0.106748, -0.801709, -2.802374, -1.108306, 1.570796, 1.677544],accel_mss,speed_ms,0,blend_radius_m)
  movel([0.107496, -0.802631, -2.802220, -1.107538, 1.570796, 1.678292],accel_mss,speed_ms,0,blend_radius_m)
  movel([0.107985, -0.804180, -2.801960, -1.106249, 1.570796, 1.678781],accel_mss,speed_ms,0,blend_radius_m)
  movel([0.108380, -0.807318, -2.801430, -1.103640, 1.570796, 1.679177],accel_mss,speed_ms,0,blend_radius_m)
  movel([0.108432, -0.810641, -2.800864, -1.100885, 1.570796, 1.679228],accel_mss,speed_ms,0,blend_radius_m)
  movel([0.108163, -0.814120, -2.800264, -1.098005, 1.570796, 1.678960],accel_mss,speed_ms,0,blend_radius_m)
  movel([0.107597, -0.817745, -2.799633, -1.095011, 1.570796, 1.678393],accel_mss,speed_ms,0,blend_radius_m)
  movel([0.106747, -0.821486, -2.798974, -1.091928, 1.570796, 1.677543],accel_mss,speed_ms,0,blend_radius_m)
  movel([0.105636, -0.825329, -2.798289, -1.088770, 1.570796, 1.676432],accel_mss,speed_ms,0,blend_radius_m)
  movel([0.104281, -0.829257, -2.797582, -1.085551, 1.570796, 1.675078],accel_mss,speed_ms,0,blend_radius_m)
  movel([0.102705, -0.833250, -2.796853, -1.082286, 1.570796, 1.673502],accel_mss,speed_ms,0,blend_radius_m)
  movel([0.098963, -0.841356, -2.795349, -1.075685, 1.570796, 1.669759],accel_mss,speed_ms,0,blend_radius_m)
  movel([0.094548, -0.849524, -2.793795, -1.069070, 1.570796, 1.665345],accel_mss,speed_ms,0,blend_radius_m)
  movel([0.089597, -0.857629, -2.792217, -1.062543, 1.570796, 1.660394],accel_mss,speed_ms,0,blend_radius_m)
  movel([0.084252, -0.865550, -2.790639, -1.056200, 1.570796, 1.655048],accel_mss,speed_ms,0,blend_radius_m)
  movel([0.071998, -0.882771, -2.787081, -1.042537, 1.570796, 1.642794],accel_mss,speed_ms,0,blend_radius_m)
  movel([0.065571, -0.891110, -2.785295, -1.035984, 1.570796, 1.636367],accel_mss,speed_ms,0,blend_radius_m)
  movel([0.062299, -0.895012, -2.784445, -1.032932, 1.570796, 1.633095],accel_mss,speed_ms,0,blend_radius_m)
  movel([0.058990, -0.898667, -2.783640, -1.030082, 1.570796, 1.629786],accel_mss,speed_ms,0,blend_radius_m)
  movel([0.056838, -0.900840, -2.783158, -1.028391, 1.570796, 1.627635],accel_mss,speed_ms,0,blend_radius_m)
  movel([0.054684, -0.902802, -2.782720, -1.026867, 1.570796, 1.625481],accel_mss,speed_ms,0,blend_radius_m)
  movel([0.052541, -0.904522, -2.782334, -1.025533, 1.570796, 1.623337],accel_mss,speed_ms,0,blend_radius_m)
  movel([0.050425, -0.905968, -2.782008, -1.024413, 1.570796, 1.621221],accel_mss,speed_ms,0,blend_radius_m)
  movel([0.048357, -0.907106, -2.781751, -1.023532, 1.570796, 1.619154],accel_mss,speed_ms,0,blend_radius_m)
  movel([0.046350, -0.907908, -2.781569, -1.022912, 1.570796, 1.617147],accel_mss,speed_ms,0,blend_radius_m)
  movel([0.044425, -0.908331, -2.781473, -1.022585, 1.570796, 1.615221],accel_mss,speed_ms,0,blend_radius_m)
  movel([0.042592, -0.908344, -2.781470, -1.022575, 1.570796, 1.613389],accel_mss,speed_ms,0,blend_radius_m)
  movel([0.040937, -0.907913, -2.781568, -1.022908, 1.570796, 1.611733],accel_mss,speed_ms,0,blend_radius_m)
  movel([0.039563, -0.907122, -2.781747, -1.023520, 1.570796, 1.610360],accel_mss,speed_ms,0,blend_radius_m)
  movel([0.034961, -0.902728, -2.782737, -1.026924, 1.570796, 1.605758],accel_mss,speed_ms,0,blend_radius_m)
  movel([0.033548, -0.901928, -2.782916, -1.027546, 1.570796, 1.604344],accel_mss,speed_ms,0,blend_radius_m)
  movel([0.031832, -0.901497, -2.783012, -1.027881, 1.570796, 1.602629],accel_mss,speed_ms,0,blend_radius_m)
  movel([0.031048, -0.901604, -2.782988, -1.027797, 1.570796, 1.601844],accel_mss,speed_ms,0,blend_radius_m)
  movel([0.030681, -0.902111, -2.782875, -1.027404, 1.570796, 1.601477],accel_mss,speed_ms,0,blend_radius_m)
  movel([0.030199, -0.903270, -2.782615, -1.026503, 1.570796, 1.600996],accel_mss,speed_ms,0,blend_radius_m)
  movel([0.028942, -0.907208, -2.781728, -1.023453, 1.570796, 1.599739],accel_mss,speed_ms,0,blend_radius_m)
  movel([0.025811, -0.918942, -2.779026, -1.014421, 1.570796, 1.596608],accel_mss,speed_ms,0,blend_radius_m)
  movel([0.020960, -0.938262, -2.774384, -0.999742, 1.570796, 1.591756],accel_mss,speed_ms,0,blend_radius_m)
  movel([0.017470, -0.948592, -2.771802, -0.991995, 1.570796, 1.588266],accel_mss,speed_ms,0,blend_radius_m)
  movel([0.013608, -0.958884, -2.769157, -0.984348, 1.570796, 1.584404],accel_mss,speed_ms,0,blend_radius_m)
  movel([0.009426, -0.969108, -2.766457, -0.976824, 1.570796, 1.580223],accel_mss,speed_ms,0,blend_radius_m)
  movel([0.004989, -0.979222, -2.763714, -0.969453, 1.570796, 1.575785],accel_mss,speed_ms,0,blend_radius_m)
  movel([-0.000886, -0.991999, -2.760143, -0.960247, 1.570796, 1.569910],accel_mss,speed_ms,0,blend_radius_m)
  movel([-0.006924, -1.004608, -2.756501, -0.951280, 1.570796, 1.563873],accel_mss,speed_ms,0,blend_radius_m)
  movel([-0.013170, -1.017002, -2.752804, -0.942583, 1.570796, 1.557626],accel_mss,speed_ms,0,blend_radius_m)
  movel([-0.019682, -1.029140, -2.749069, -0.934180, 1.570796, 1.551114],accel_mss,speed_ms,0,blend_radius_m)
  movel([-0.026507, -1.040975, -2.745314, -0.926100, 1.570796, 1.544290],accel_mss,speed_ms,0,blend_radius_m)
  movel([-0.030048, -1.046767, -2.743435, -0.922187, 1.570796, 1.540749],accel_mss,speed_ms,0,blend_radius_m)
  movel([-0.033689, -1.052474, -2.741557, -0.918359, 1.570796, 1.537107],accel_mss,speed_ms,0,blend_radius_m)
  movel([-0.037435, -1.058089, -2.739682, -0.914618, 1.570796, 1.533362],accel_mss,speed_ms,0,blend_radius_m)
  movel([-0.041287, -1.063604, -2.737815, -0.910970, 1.570796, 1.529509],accel_mss,speed_ms,0,blend_radius_m)
  movel([-0.045255, -1.069024, -2.735955, -0.907410, 1.570796, 1.525541],accel_mss,speed_ms,0,blend_radius_m)
  movel([-0.049349, -1.074339, -2.734107, -0.903943, 1.570796, 1.521448],accel_mss,speed_ms,0,blend_radius_m)
  movel([-0.054352, -1.080512, -2.731930, -0.899948, 1.570796, 1.516444],accel_mss,speed_ms,0,blend_radius_m)
  movel([-0.056958, -1.083475, -2.730873, -0.898041, 1.570796, 1.513838],accel_mss,speed_ms,0,blend_radius_m)
  movel([-0.061649, -1.088234, -2.729159, -0.894996, 1.570796, 1.509147],accel_mss,speed_ms,0,blend_radius_m)
  movel([-0.064077, -1.090406, -2.728370, -0.893613, 1.570796, 1.506719],accel_mss,speed_ms,0,blend_radius_m)
  movel([-0.066519, -1.092141, -2.727736, -0.892511, 1.570796, 1.504277],accel_mss,speed_ms,0,blend_radius_m)
  movel([-0.067609, -1.092635, -2.727556, -0.892198, 1.570796, 1.503188],accel_mss,speed_ms,0,blend_radius_m)
  movel([-0.068545, -1.092774, -2.727505, -0.892110, 1.570796, 1.502251],accel_mss,speed_ms,0,blend_radius_m)
  movel([-0.067892, -1.090183, -2.728451, -0.893755, 1.570796, 1.502904],accel_mss,speed_ms,0,blend_radius_m)
  movel([-0.067596, -1.087727, -2.729342, -0.895320, 1.570796, 1.503200],accel_mss,speed_ms,0,blend_radius_m)
  movel([-0.067673, -1.086667, -2.729725, -0.895997, 1.570796, 1.503124],accel_mss,speed_ms,0,blend_radius_m)
  movel([-0.067948, -1.085783, -2.730044, -0.896562, 1.570796, 1.502849],accel_mss,speed_ms,0,blend_radius_m)
  movel([-0.068456, -1.085118, -2.730283, -0.896988, 1.570796, 1.502340],accel_mss,speed_ms,0,blend_radius_m)
  movel([-0.069242, -1.084730, -2.730423, -0.897236, 1.570796, 1.501554],accel_mss,speed_ms,0,blend_radius_m)
  movel([-0.071652, -1.084503, -2.730504, -0.897382, 1.570796, 1.499145],accel_mss,speed_ms,0,blend_radius_m)
  movel([-0.072322, -1.084160, -2.730627, -0.897602, 1.570796, 1.498475],accel_mss,speed_ms,0,blend_radius_m)
  movel([-0.072785, -1.083602, -2.730827, -0.897960, 1.570796, 1.498011],accel_mss,speed_ms,0,blend_radius_m)
  movel([-0.073179, -1.081983, -2.731406, -0.899000, 1.570796, 1.497617],accel_mss,speed_ms,0,blend_radius_m)
  movel([-0.073051, -1.079928, -2.732137, -0.900324, 1.570796, 1.497746],accel_mss,speed_ms,0,blend_radius_m)
  movel([-0.072608, -1.077725, -2.732917, -0.901747, 1.570796, 1.498188],accel_mss,speed_ms,0,blend_radius_m)
  movel([-0.070858, -1.070937, -2.735293, -0.906159, 1.570796, 1.499938],accel_mss,speed_ms,0,blend_radius_m)
  movel([-0.068698, -1.063915, -2.737709, -0.910765, 1.570796, 1.502098],accel_mss,speed_ms,0,blend_radius_m)
  movel([-0.067395, -1.060333, -2.738926, -0.913131, 1.570796, 1.503402],accel_mss,speed_ms,0,blend_radius_m)
  movel([-0.065910, -1.056707, -2.740146, -0.915536, 1.570796, 1.504886],accel_mss,speed_ms,0,blend_radius_m)
  movel([-0.064215, -1.053048, -2.741366, -0.917975, 1.570796, 1.506582],accel_mss,speed_ms,0,blend_radius_m)
  movel([-0.062279, -1.049360, -2.742585, -0.920444, 1.570796, 1.508517],accel_mss,speed_ms,0,blend_radius_m)
  movel([-0.060072, -1.045797, -2.743751, -0.922841, 1.570796, 1.510725],accel_mss,speed_ms,0,blend_radius_m)
  movel([-0.052653, -1.035496, -2.747066, -0.929827, 1.570796, 1.518143],accel_mss,speed_ms,0,blend_radius_m)
  movel([-0.046893, -1.026534, -2.749880, -0.935974, 1.570796, 1.523903],accel_mss,speed_ms,0,blend_radius_m)
  movel([-0.041269, -1.017369, -2.752693, -0.942327, 1.570796, 1.529527],accel_mss,speed_ms,0,blend_radius_m)
  movel([-0.038775, -1.013190, -2.753954, -0.945245, 1.570796, 1.532021],accel_mss,speed_ms,0,blend_radius_m)
  speed_ms = 0.005
  movel([-0.038775, -1.003253, -2.748331, -0.960805, 1.570796, 1.532021],accel_mss,speed_ms,0,blend_radius_m)
  speed_ms = 0.040
  movel([-0.089816, -1.077062, -2.724259, -0.911067, 1.570796, 1.480980],accel_mss,speed_ms,0,blend_radius_m)
  speed_ms = 0.005
  movel([-0.089816, -1.087093, -2.729571, -0.895724, 1.570796, 1.480980],accel_mss,speed_ms,0,blend_radius_m)
  speed_ms = 0.025
  movel([-0.085381, -1.090136, -2.728468, -0.893785, 1.570796, 1.485415],accel_mss,speed_ms,0,blend_radius_m)
  movel([-0.083192, -1.091957, -2.727804, -0.892628, 1.570796, 1.487604],accel_mss,speed_ms,0,blend_radius_m)
  movel([-0.081191, -1.094019, -2.727048, -0.891322, 1.570796, 1.489606],accel_mss,speed_ms,0,blend_radius_m)
  movel([-0.079489, -1.096337, -2.726194, -0.889858, 1.570796, 1.491307],accel_mss,speed_ms,0,blend_radius_m)
  movel([-0.078209, -1.098931, -2.725232, -0.888226, 1.570796, 1.492587],accel_mss,speed_ms,0,blend_radius_m)
  movel([-0.077467, -1.101824, -2.724153, -0.886413, 1.570796, 1.493329],accel_mss,speed_ms,0,blend_radius_m)
  movel([-0.077335, -1.103390, -2.723565, -0.885434, 1.570796, 1.493461],accel_mss,speed_ms,0,blend_radius_m)
  movel([-0.077380, -1.105033, -2.722946, -0.884410, 1.570796, 1.493416],accel_mss,speed_ms,0,blend_radius_m)
  movel([-0.078452, -1.104725, -2.723062, -0.884602, 1.570796, 1.492345],accel_mss,speed_ms,0,blend_radius_m)
  movel([-0.079150, -1.104138, -2.723283, -0.884967, 1.570796, 1.491646],accel_mss,speed_ms,0,blend_radius_m)
  movel([-0.080624, -1.102732, -2.723812, -0.885845, 1.570796, 1.490172],accel_mss,speed_ms,0,blend_radius_m)
  movel([-0.082650, -1.101733, -2.724187, -0.886469, 1.570796, 1.488147],accel_mss,speed_ms,0,blend_radius_m)
  movel([-0.084885, -1.101010, -2.724457, -0.886922, 1.570796, 1.485911],accel_mss,speed_ms,0,blend_radius_m)
  movel([-0.087305, -1.100550, -2.724629, -0.887210, 1.570796, 1.483491],accel_mss,speed_ms,0,blend_radius_m)
  movel([-0.089883, -1.100347, -2.724705, -0.887337, 1.570796, 1.480913],accel_mss,speed_ms,0,blend_radius_m)
  movel([-0.092594, -1.100390, -2.724689, -0.887311, 1.570796, 1.478203],accel_mss,speed_ms,0,blend_radius_m)
  movel([-0.095409, -1.100671, -2.724584, -0.887134, 1.570796, 1.475387],accel_mss,speed_ms,0,blend_radius_m)
  movel([-0.098307, -1.101183, -2.724393, -0.886814, 1.570796, 1.472490],accel_mss,speed_ms,0,blend_radius_m)
  movel([-0.101256, -1.101910, -2.724120, -0.886358, 1.570796, 1.469540],accel_mss,speed_ms,0,blend_radius_m)
  movel([-0.103243, -1.102563, -2.723876, -0.885950, 1.570796, 1.467553],accel_mss,speed_ms,0,blend_radius_m)
  movel([-0.104813, -1.103279, -2.723607, -0.885504, 1.570796, 1.465983],accel_mss,speed_ms,0,blend_radius_m)
  movel([-0.105996, -1.104044, -2.723319, -0.885026, 1.570796, 1.464800],accel_mss,speed_ms,0,blend_radius_m)
  movel([-0.106828, -1.104848, -2.723016, -0.884525, 1.570796, 1.463969],accel_mss,speed_ms,0,blend_radius_m)
  movel([-0.107346, -1.105690, -2.722698, -0.884001, 1.570796, 1.463451],accel_mss,speed_ms,0,blend_radius_m)
  movel([-0.107582, -1.106558, -2.722369, -0.883462, 1.570796, 1.463214],accel_mss,speed_ms,0,blend_radius_m)
  movel([-0.107579, -1.107447, -2.722032, -0.882910, 1.570796, 1.463218],accel_mss,speed_ms,0,blend_radius_m)
  movel([-0.107365, -1.108347, -2.721690, -0.882352, 1.570796, 1.463432],accel_mss,speed_ms,0,blend_radius_m)
  movel([-0.106462, -1.110164, -2.720997, -0.881228, 1.570796, 1.464334],accel_mss,speed_ms,0,blend_radius_m)
  movel([-0.102469, -1.115261, -2.719037, -0.878092, 1.570796, 1.468328],accel_mss,speed_ms,0,blend_radius_m)
  movel([-0.105068, -1.114356, -2.719386, -0.878647, 1.570796, 1.465728],accel_mss,speed_ms,0,blend_radius_m)
  movel([-0.110164, -1.112418, -2.720133, -0.879838, 1.570796, 1.460632],accel_mss,speed_ms,0,blend_radius_m)
  movel([-0.113027, -1.111934, -2.720319, -0.880136, 1.570796, 1.457770],accel_mss,speed_ms,0,blend_radius_m)
  movel([-0.116461, -1.111871, -2.720343, -0.880175, 1.570796, 1.454335],accel_mss,speed_ms,0,blend_radius_m)
  movel([-0.120018, -1.112021, -2.720286, -0.880083, 1.570796, 1.450778],accel_mss,speed_ms,0,blend_radius_m)
  movel([-0.127213, -1.112491, -2.720105, -0.879793, 1.570796, 1.443583],accel_mss,speed_ms,0,blend_radius_m)
  movel([-0.130713, -1.112583, -2.720069, -0.879736, 1.570796, 1.440083],accel_mss,speed_ms,0,blend_radius_m)
  movel([-0.134055, -1.112426, -2.720130, -0.879833, 1.570796, 1.436742],accel_mss,speed_ms,0,blend_radius_m)
  movel([-0.137170, -1.111909, -2.720329, -0.880152, 1.570796, 1.433626],accel_mss,speed_ms,0,blend_radius_m)
  movel([-0.139995, -1.110910, -2.720711, -0.880767, 1.570796, 1.430802],accel_mss,speed_ms,0,blend_radius_m)
  movel([-0.137192, -1.115418, -2.718976, -0.877995, 1.570796, 1.433605],accel_mss,speed_ms,0,blend_radius_m)
  movel([-0.135602, -1.117594, -2.718131, -0.876664, 1.570796, 1.435194],accel_mss,speed_ms,0,blend_radius_m)
  movel([-0.133826, -1.119315, -2.717460, -0.875614, 1.570796, 1.436971],accel_mss,speed_ms,0,blend_radius_m)
  movel([-0.136672, -1.118444, -2.717800, -0.876145, 1.570796, 1.434124],accel_mss,speed_ms,0,blend_radius_m)
  movel([-0.139763, -1.117945, -2.717994, -0.876449, 1.570796, 1.431033],accel_mss,speed_ms,0,blend_radius_m)
  movel([-0.146189, -1.117328, -2.718235, -0.876827, 1.570796, 1.424608],accel_mss,speed_ms,0,blend_radius_m)
  movel([-0.148233, -1.116943, -2.718384, -0.877062, 1.570796, 1.422563],accel_mss,speed_ms,0,blend_radius_m)
  movel([-0.150068, -1.116334, -2.718621, -0.877434, 1.570796, 1.420728],accel_mss,speed_ms,0,blend_radius_m)
  movel([-0.153333, -1.114665, -2.719267, -0.878457, 1.570796, 1.417463],accel_mss,speed_ms,0,blend_radius_m)
  movel([-0.156453, -1.112786, -2.719991, -0.879611, 1.570796, 1.414344],accel_mss,speed_ms,0,blend_radius_m)
  movel([-0.159894, -1.111176, -2.720609, -0.880603, 1.570796, 1.410903],accel_mss,speed_ms,0,blend_radius_m)
  movel([-0.161112, -1.110847, -2.720736, -0.880806, 1.570796, 1.409685],accel_mss,speed_ms,0,blend_radius_m)
  movel([-0.162467, -1.110751, -2.720773, -0.880866, 1.570796, 1.408329],accel_mss,speed_ms,0,blend_radius_m)
  movel([-0.163937, -1.111036, -2.720663, -0.880690, 1.570796, 1.406859],accel_mss,speed_ms,0,blend_radius_m)
  movel([-0.164701, -1.111362, -2.720538, -0.880489, 1.570796, 1.406095],accel_mss,speed_ms,0,blend_radius_m)
  movel([-0.165483, -1.111841, -2.720355, -0.880194, 1.570796, 1.405313],accel_mss,speed_ms,0,blend_radius_m)
  movel([-0.166307, -1.112511, -2.720097, -0.879781, 1.570796, 1.404490],accel_mss,speed_ms,0,blend_radius_m)
  movel([-0.167031, -1.113275, -2.719803, -0.879311, 1.570796, 1.403765],accel_mss,speed_ms,0,blend_radius_m)
  movel([-0.168230, -1.115010, -2.719133, -0.878245, 1.570796, 1.402566],accel_mss,speed_ms,0,blend_radius_m)
  movel([-0.169139, -1.116883, -2.718408, -0.877098, 1.570796, 1.401658],accel_mss,speed_ms,0,blend_radius_m)
  movel([-0.169815, -1.118729, -2.717689, -0.875971, 1.570796, 1.400982],accel_mss,speed_ms,0,blend_radius_m)
  movel([-0.170869, -1.116461, -2.718571, -0.877357, 1.570796, 1.399927],accel_mss,speed_ms,0,blend_radius_m)
  movel([-0.172146, -1.114433, -2.719357, -0.878600, 1.570796, 1.398650],accel_mss,speed_ms,0,blend_radius_m)
  movel([-0.175130, -1.110853, -2.720733, -0.880803, 1.570796, 1.395666],accel_mss,speed_ms,0,blend_radius_m)
  movel([-0.178288, -1.107452, -2.722030, -0.882907, 1.570796, 1.392508],accel_mss,speed_ms,0,blend_radius_m)
  movel([-0.181130, -1.103672, -2.723459, -0.885258, 1.570796, 1.389666],accel_mss,speed_ms,0,blend_radius_m)
  movel([-0.181947, -1.101943, -2.724108, -0.886338, 1.570796, 1.388849],accel_mss,speed_ms,0,blend_radius_m)
  movel([-0.182498, -1.099942, -2.724856, -0.887591, 1.570796, 1.388298],accel_mss,speed_ms,0,blend_radius_m)
  movel([-0.182819, -1.097720, -2.725682, -0.888987, 1.570796, 1.387977],accel_mss,speed_ms,0,blend_radius_m)
  movel([-0.182952, -1.095341, -2.726561, -0.890486, 1.570796, 1.387845],accel_mss,speed_ms,0,blend_radius_m)
  movel([-0.182776, -1.090309, -2.728405, -0.893675, 1.570796, 1.388020],accel_mss,speed_ms,0,blend_radius_m)
  movel([-0.182269, -1.085305, -2.730216, -0.896868, 1.570796, 1.388528],accel_mss,speed_ms,0,blend_radius_m)
  speed_ms = 0.005
  movel([-0.182269, -1.075274, -2.724896, -0.912219, 1.570796, 1.388528],accel_mss,speed_ms,0,blend_radius_m)
  speed_ms = 0.040
  # Splitting Linear movement in 2 (instruction 806: MoveL 765)
  movel([-0.154336, -1.000413, -2.749171, -0.962805, 1.570796, 1.416460],accel_mss,speed_ms,0,blend_radius_m)
  movel([-0.121695, -0.915912, -2.771520, -1.024957, 1.570796, 1.449101],accel_mss,speed_ms,0,blend_radius_m)
  speed_ms = 0.005
  movel([-0.121695, -0.925478, -2.777483, -1.009429, 1.570796, 1.449101],accel_mss,speed_ms,0,blend_radius_m)
  speed_ms = 0.025
  movel([-0.123729, -0.928016, -2.776876, -1.007497, 1.570796, 1.447067],accel_mss,speed_ms,0,blend_radius_m)
  movel([-0.123869, -0.928434, -2.776776, -1.007179, 1.570796, 1.446928],accel_mss,speed_ms,0,blend_radius_m)
  movel([-0.123677, -0.928895, -2.776665, -1.006829, 1.570796, 1.447119],accel_mss,speed_ms,0,blend_radius_m)
  movel([-0.122387, -0.929956, -2.776410, -1.006023, 1.570796, 1.448409],accel_mss,speed_ms,0,blend_radius_m)
  movel([-0.116786, -0.932544, -2.775783, -1.004061, 1.570796, 1.454011],accel_mss,speed_ms,0,blend_radius_m)
  movel([-0.108296, -0.935614, -2.775035, -1.001740, 1.570796, 1.462501],accel_mss,speed_ms,0,blend_radius_m)
  movel([-0.098262, -0.938973, -2.774209, -0.999207, 1.570796, 1.472535],accel_mss,speed_ms,0,blend_radius_m)
  movel([-0.078691, -0.945470, -2.772590, -0.994329, 1.570796, 1.492105],accel_mss,speed_ms,0,blend_radius_m)
  movel([-0.067694, -0.949059, -2.771683, -0.991646, 1.570796, 1.503103],accel_mss,speed_ms,0,blend_radius_m)
  movel([-0.066628, -0.949228, -2.771640, -0.991520, 1.570796, 1.504168],accel_mss,speed_ms,0,blend_radius_m)
  movel([-0.065426, -0.949141, -2.771662, -0.991585, 1.570796, 1.505370],accel_mss,speed_ms,0,blend_radius_m)
  movel([-0.064169, -0.948645, -2.771789, -0.991956, 1.570796, 1.506628],accel_mss,speed_ms,0,blend_radius_m)
  movel([-0.063539, -0.948197, -2.771902, -0.992290, 1.570796, 1.507257],accel_mss,speed_ms,0,blend_radius_m)
  movel([-0.062925, -0.947587, -2.772056, -0.992746, 1.570796, 1.507871],accel_mss,speed_ms,0,blend_radius_m)
  movel([-0.062039, -0.946272, -2.772388, -0.993729, 1.570796, 1.508758],accel_mss,speed_ms,0,blend_radius_m)
  movel([-0.061407, -0.944895, -2.772734, -0.994759, 1.570796, 1.509389],accel_mss,speed_ms,0,blend_radius_m)
  movel([-0.058516, -0.937255, -2.774633, -1.000502, 1.570796, 1.512280],accel_mss,speed_ms,0,blend_radius_m)
  movel([-0.056125, -0.929684, -2.776475, -1.006230, 1.570796, 1.514671],accel_mss,speed_ms,0,blend_radius_m)
  movel([-0.054216, -0.922220, -2.778255, -1.011914, 1.570796, 1.516580],accel_mss,speed_ms,0,blend_radius_m)
  movel([-0.052750, -0.914889, -2.779969, -1.017531, 1.570796, 1.518046],accel_mss,speed_ms,0,blend_radius_m)
  movel([-0.051705, -0.907721, -2.781611, -1.023056, 1.570796, 1.519091],accel_mss,speed_ms,0,blend_radius_m)
  movel([-0.051044, -0.900744, -2.783179, -1.028466, 1.570796, 1.519752],accel_mss,speed_ms,0,blend_radius_m)
  movel([-0.050737, -0.893988, -2.784669, -1.033732, 1.570796, 1.520059],accel_mss,speed_ms,0,blend_radius_m)
  movel([-0.050750, -0.887488, -2.786076, -1.038825, 1.570796, 1.520046],accel_mss,speed_ms,0,blend_radius_m)
  movel([-0.050960, -0.884671, -2.786678, -1.041040, 1.570796, 1.519836],accel_mss,speed_ms,0,blend_radius_m)
  movel([-0.051433, -0.882235, -2.787194, -1.042960, 1.570796, 1.519363],accel_mss,speed_ms,0,blend_radius_m)
  movel([-0.052166, -0.880177, -2.787628, -1.044584, 1.570796, 1.518631],accel_mss,speed_ms,0,blend_radius_m)
  movel([-0.053142, -0.878484, -2.787983, -1.045922, 1.570796, 1.517655],accel_mss,speed_ms,0,blend_radius_m)
  movel([-0.054358, -0.877156, -2.788260, -1.046973, 1.570796, 1.516439],accel_mss,speed_ms,0,blend_radius_m)
  movel([-0.055805, -0.876187, -2.788462, -1.047740, 1.570796, 1.514992],accel_mss,speed_ms,0,blend_radius_m)
  movel([-0.057470, -0.875559, -2.788592, -1.048238, 1.570796, 1.513326],accel_mss,speed_ms,0,blend_radius_m)
  movel([-0.059349, -0.875268, -2.788652, -1.048469, 1.570796, 1.511448],accel_mss,speed_ms,0,blend_radius_m)
  movel([-0.061426, -0.875305, -2.788645, -1.048440, 1.570796, 1.509370],accel_mss,speed_ms,0,blend_radius_m)
  movel([-0.063692, -0.875659, -2.788571, -1.048159, 1.570796, 1.507104],accel_mss,speed_ms,0,blend_radius_m)
  movel([-0.066142, -0.876319, -2.788434, -1.047636, 1.570796, 1.504655],accel_mss,speed_ms,0,blend_radius_m)
  movel([-0.068755, -0.877274, -2.788235, -1.046879, 1.570796, 1.502042],accel_mss,speed_ms,0,blend_radius_m)
  movel([-0.074446, -0.880029, -2.787659, -1.044701, 1.570796, 1.496350],accel_mss,speed_ms,0,blend_radius_m)
  movel([-0.080671, -0.883820, -2.786859, -1.041710, 1.570796, 1.490125],accel_mss,speed_ms,0,blend_radius_m)
  movel([-0.086258, -0.887856, -2.785997, -1.038536, 1.570796, 1.484538],accel_mss,speed_ms,0,blend_radius_m)
  movel([-0.091716, -0.892402, -2.785015, -1.034972, 1.570796, 1.479080],accel_mss,speed_ms,0,blend_radius_m)
  movel([-0.097048, -0.897380, -2.783925, -1.031084, 1.570796, 1.473748],accel_mss,speed_ms,0,blend_radius_m)
  movel([-0.102248, -0.902688, -2.782745, -1.026955, 1.570796, 1.468548],accel_mss,speed_ms,0,blend_radius_m)
  movel([-0.107307, -0.908234, -2.781495, -1.022660, 1.570796, 1.463490],accel_mss,speed_ms,0,blend_radius_m)
  movel([-0.112236, -0.913938, -2.780189, -1.018263, 1.570796, 1.458561],accel_mss,speed_ms,0,blend_radius_m)
  movel([-0.121695, -0.925478, -2.777483, -1.009429, 1.570796, 1.449101],accel_mss,speed_ms,0,blend_radius_m)
  movel([-0.123729, -0.928016, -2.776876, -1.007497, 1.570796, 1.447067],accel_mss,speed_ms,0,blend_radius_m)
  movel([-0.123869, -0.928434, -2.776776, -1.007179, 1.570796, 1.446928],accel_mss,speed_ms,0,blend_radius_m)
  movel([-0.123677, -0.928895, -2.776665, -1.006829, 1.570796, 1.447119],accel_mss,speed_ms,0,blend_radius_m)
  movel([-0.123269, -0.929232, -2.776584, -1.006573, 1.570796, 1.447527],accel_mss,speed_ms,0,blend_radius_m)
  speed_ms = 0.005
  movel([-0.123269, -0.919645, -2.770635, -1.022109, 1.570796, 1.447527],accel_mss,speed_ms,0,blend_radius_m)
  speed_ms = 0.040
  movel([-0.141809, -0.897042, -2.775859, -1.039488, 1.570796, 1.428988],accel_mss,speed_ms,0,blend_radius_m)
  speed_ms = 0.005
  movel([-0.141809, -0.906488, -2.781891, -1.024010, 1.570796, 1.428988],accel_mss,speed_ms,0,blend_radius_m)
  speed_ms = 0.025
  movel([-0.142140, -0.904068, -2.782436, -1.025884, 1.570796, 1.428656],accel_mss,speed_ms,0,blend_radius_m)
  movel([-0.142908, -0.902017, -2.782896, -1.027476, 1.570796, 1.427888],accel_mss,speed_ms,0,blend_radius_m)
  movel([-0.144096, -0.900389, -2.783258, -1.028741, 1.570796, 1.426701],accel_mss,speed_ms,0,blend_radius_m)
  movel([-0.145674, -0.899220, -2.783518, -1.029651, 1.570796, 1.425122],accel_mss,speed_ms,0,blend_radius_m)
  movel([-0.150413, -0.897523, -2.783893, -1.030973, 1.570796, 1.420383],accel_mss,speed_ms,0,blend_radius_m)
  movel([-0.151583, -0.896805, -2.784051, -1.031533, 1.570796, 1.419213],accel_mss,speed_ms,0,blend_radius_m)
  movel([-0.152432, -0.895866, -2.784258, -1.032265, 1.570796, 1.418365],accel_mss,speed_ms,0,blend_radius_m)
  movel([-0.152803, -0.894661, -2.784522, -1.033206, 1.570796, 1.417993],accel_mss,speed_ms,0,blend_radius_m)
  movel([-0.152536, -0.893128, -2.784857, -1.034404, 1.570796, 1.418260],accel_mss,speed_ms,0,blend_radius_m)
  movel([-0.151543, -0.891171, -2.785282, -1.035936, 1.570796, 1.419254],accel_mss,speed_ms,0,blend_radius_m)
  movel([-0.150265, -0.889649, -2.785611, -1.037129, 1.570796, 1.420531],accel_mss,speed_ms,0,blend_radius_m)
  movel([-0.148786, -0.888509, -2.785857, -1.038024, 1.570796, 1.422010],accel_mss,speed_ms,0,blend_radius_m)
  movel([-0.147199, -0.887699, -2.786031, -1.038659, 1.570796, 1.423597],accel_mss,speed_ms,0,blend_radius_m)
  movel([-0.144077, -0.886874, -2.786208, -1.039308, 1.570796, 1.426719],accel_mss,speed_ms,0,blend_radius_m)
  movel([-0.141608, -0.886743, -2.786236, -1.039410, 1.570796, 1.429189],accel_mss,speed_ms,0,blend_radius_m)
  movel([-0.142716, -0.884245, -2.786768, -1.041376, 1.570796, 1.428081],accel_mss,speed_ms,0,blend_radius_m)
  movel([-0.144331, -0.882355, -2.787169, -1.042865, 1.570796, 1.426465],accel_mss,speed_ms,0,blend_radius_m)
  movel([-0.148487, -0.879656, -2.787737, -1.044995, 1.570796, 1.422309],accel_mss,speed_ms,0,blend_radius_m)
  movel([-0.152861, -0.877101, -2.788272, -1.047017, 1.570796, 1.417935],accel_mss,speed_ms,0,blend_radius_m)
  movel([-0.154755, -0.875386, -2.788628, -1.048375, 1.570796, 1.416041],accel_mss,speed_ms,0,blend_radius_m)
  movel([-0.156241, -0.873108, -2.789099, -1.050182, 1.570796, 1.414555],accel_mss,speed_ms,0,blend_radius_m)
  movel([-0.156900, -0.871384, -2.789453, -1.051552, 1.570796, 1.413896],accel_mss,speed_ms,0,blend_radius_m)
  movel([-0.157213, -0.869787, -2.789779, -1.052822, 1.570796, 1.413584],accel_mss,speed_ms,0,blend_radius_m)
  movel([-0.157211, -0.868322, -2.790078, -1.053989, 1.570796, 1.413585],accel_mss,speed_ms,0,blend_radius_m)
  movel([-0.156924, -0.866997, -2.790346, -1.055046, 1.570796, 1.413873],accel_mss,speed_ms,0,blend_radius_m)
  movel([-0.156395, -0.865826, -2.790583, -1.055980, 1.570796, 1.414402],accel_mss,speed_ms,0,blend_radius_m)
  movel([-0.155651, -0.864803, -2.790789, -1.056797, 1.570796, 1.415145],accel_mss,speed_ms,0,blend_radius_m)
  movel([-0.154736, -0.863947, -2.790961, -1.057481, 1.570796, 1.416060],accel_mss,speed_ms,0,blend_radius_m)
  movel([-0.153677, -0.863259, -2.791099, -1.058031, 1.570796, 1.417119],accel_mss,speed_ms,0,blend_radius_m)
  movel([-0.152514, -0.862752, -2.791200, -1.058437, 1.570796, 1.418282],accel_mss,speed_ms,0,blend_radius_m)
  movel([-0.151289, -0.862435, -2.791264, -1.058691, 1.570796, 1.419507],accel_mss,speed_ms,0,blend_radius_m)
  movel([-0.148777, -0.862389, -2.791273, -1.058727, 1.570796, 1.422019],accel_mss,speed_ms,0,blend_radius_m)
  movel([-0.146432, -0.863178, -2.791115, -1.058096, 1.570796, 1.424365],accel_mss,speed_ms,0,blend_radius_m)
  movel([-0.144538, -0.864858, -2.790778, -1.056753, 1.570796, 1.426258],accel_mss,speed_ms,0,blend_radius_m)
  movel([-0.144291, -0.861792, -2.791392, -1.059205, 1.570796, 1.426505],accel_mss,speed_ms,0,blend_radius_m)
  movel([-0.144419, -0.859148, -2.791917, -1.061324, 1.570796, 1.426377],accel_mss,speed_ms,0,blend_radius_m)
  movel([-0.144844, -0.856835, -2.792373, -1.063180, 1.570796, 1.425952],accel_mss,speed_ms,0,blend_radius_m)
  movel([-0.147033, -0.850767, -2.793556, -1.068066, 1.570796, 1.423764],accel_mss,speed_ms,0,blend_radius_m)
  movel([-0.148397, -0.846354, -2.794403, -1.071633, 1.570796, 1.422399],accel_mss,speed_ms,0,blend_radius_m)
  movel([-0.148692, -0.844295, -2.794794, -1.073300, 1.570796, 1.422104],accel_mss,speed_ms,0,blend_radius_m)
  movel([-0.148704, -0.842320, -2.795167, -1.074902, 1.570796, 1.422092],accel_mss,speed_ms,0,blend_radius_m)
  movel([-0.148469, -0.840458, -2.795517, -1.076414, 1.570796, 1.422328],accel_mss,speed_ms,0,blend_radius_m)
  movel([-0.148012, -0.838730, -2.795840, -1.077819, 1.570796, 1.422784],accel_mss,speed_ms,0,blend_radius_m)
  movel([-0.147373, -0.837162, -2.796132, -1.079095, 1.570796, 1.423424],accel_mss,speed_ms,0,blend_radius_m)
  movel([-0.146578, -0.835775, -2.796388, -1.080225, 1.570796, 1.424218],accel_mss,speed_ms,0,blend_radius_m)
  movel([-0.145663, -0.834595, -2.796606, -1.081187, 1.570796, 1.425134],accel_mss,speed_ms,0,blend_radius_m)
  movel([-0.144659, -0.833649, -2.796780, -1.081960, 1.570796, 1.426137],accel_mss,speed_ms,0,blend_radius_m)
  movel([-0.143601, -0.832961, -2.796906, -1.082521, 1.570796, 1.427195],accel_mss,speed_ms,0,blend_radius_m)
  movel([-0.142525, -0.832555, -2.796981, -1.082853, 1.570796, 1.428271],accel_mss,speed_ms,0,blend_radius_m)
  movel([-0.141459, -0.832453, -2.796999, -1.082936, 1.570796, 1.429337],accel_mss,speed_ms,0,blend_radius_m)
  movel([-0.140438, -0.832684, -2.796957, -1.082748, 1.570796, 1.430358],accel_mss,speed_ms,0,blend_radius_m)
  movel([-0.139501, -0.833273, -2.796849, -1.082267, 1.570796, 1.431295],accel_mss,speed_ms,0,blend_radius_m)
  movel([-0.138678, -0.834240, -2.796672, -1.081478, 1.570796, 1.432119],accel_mss,speed_ms,0,blend_radius_m)
  movel([-0.138001, -0.835609, -2.796419, -1.080361, 1.570796, 1.432795],accel_mss,speed_ms,0,blend_radius_m)
  movel([-0.137501, -0.837395, -2.796088, -1.078906, 1.570796, 1.433296],accel_mss,speed_ms,0,blend_radius_m)
  movel([-0.136094, -0.834132, -2.796691, -1.081565, 1.570796, 1.434702],accel_mss,speed_ms,0,blend_radius_m)
  movel([-0.135009, -0.830995, -2.797266, -1.084128, 1.570796, 1.435788],accel_mss,speed_ms,0,blend_radius_m)
  movel([-0.134183, -0.827959, -2.797817, -1.086614, 1.570796, 1.436613],accel_mss,speed_ms,0,blend_radius_m)
  movel([-0.133548, -0.824994, -2.798349, -1.089045, 1.570796, 1.437248],accel_mss,speed_ms,0,blend_radius_m)
  movel([-0.131530, -0.813318, -2.800403, -1.098668, 1.570796, 1.439266],accel_mss,speed_ms,0,blend_radius_m)
  movel([-0.130668, -0.808935, -2.801155, -1.102299, 1.570796, 1.440128],accel_mss,speed_ms,0,blend_radius_m)
  movel([-0.129218, -0.803528, -2.802070, -1.106792, 1.570796, 1.441578],accel_mss,speed_ms,0,blend_radius_m)
  movel([-0.128102, -0.800765, -2.802531, -1.109093, 1.570796, 1.442695],accel_mss,speed_ms,0,blend_radius_m)
  movel([-0.126634, -0.798146, -2.802965, -1.111278, 1.570796, 1.444162],accel_mss,speed_ms,0,blend_radius_m)
  movel([-0.125742, -0.796928, -2.803165, -1.112296, 1.570796, 1.445055],accel_mss,speed_ms,0,blend_radius_m)
  movel([-0.123614, -0.794765, -2.803519, -1.114105, 1.570796, 1.447182],accel_mss,speed_ms,0,blend_radius_m)
  movel([-0.122358, -0.793858, -2.803667, -1.114864, 1.570796, 1.448438],accel_mss,speed_ms,0,blend_radius_m)
